(* IEC 61131-3 sources: plcassist-cli/packages/volt-lsp-iec/test-corpus/pro2193/Device/Plc Logic/Application/09 Misc/Library Manager/L_TT1P_TechnologyModules, 210 files *)

(* ---- L_MB1P_CONSTANTS.gvl ---- *)
VAR_GLOBAL
	GC_DWCHECKIDTAPPETREF : DWORD := 16#DC34;
	GC_LREPSILON : LREAL := 1E-06;
	GC_POSITIVE_LIMIT_32BIT : LREAL := 2147483647;
	GC_NEGATIVE_LIMIT_32BIT : LREAL := -2147483647;
	GC_PI : LREAL := 3.1415926535897931;
END_VAR

(* ---- L_MB1P_GLOBAL.gvl ---- *)
VAR_GLOBAL
END_VAR

(* ---- ITF_DATABUS.itf ---- *)
INTERFACE ITF_DATABUS
END_INTERFACE

(* ---- ITF_DATABUSPAR.itf ---- *)
INTERFACE ITF_DATABUSPAR
END_INTERFACE

(* ---- ITF_LIST.itf ---- *)
INTERFACE ITF_LIST
END_INTERFACE

(* ---- GETBOOLEANPROPERTY.fun ---- *)
FUNCTION GETBOOLEANPROPERTY : BOOL
VAR_INPUT
	STKEY : WSTRING;
END_VAR
END_FUNCTION

(* ---- GETCOMPANY.fun ---- *)
FUNCTION GETCOMPANY : WSTRING
END_FUNCTION

(* ---- GETNUMBERPROPERTY.fun ---- *)
FUNCTION GETNUMBERPROPERTY : DINT
VAR_INPUT
	STKEY : WSTRING;
END_VAR
END_FUNCTION

(* ---- GETTEXTPROPERTY.fun ---- *)
FUNCTION GETTEXTPROPERTY : WSTRING
VAR_INPUT
	STKEY : WSTRING;
END_VAR
END_FUNCTION

(* ---- GETTEXTPROPERTY2.fun ---- *)
FUNCTION GETTEXTPROPERTY2 : POINTER TO WSTRING
VAR_INPUT
	STKEY : WSTRING;
END_VAR
END_FUNCTION

(* ---- GETTITLE.fun ---- *)
FUNCTION GETTITLE : WSTRING
END_FUNCTION

(* ---- GETVERSION.fun ---- *)
FUNCTION GETVERSION : VERSION
END_FUNCTION

(* ---- GETVERSIONPROPERTY.fun ---- *)
FUNCTION GETVERSIONPROPERTY : VERSION
VAR_INPUT
	STKEY : WSTRING;
END_VAR
END_FUNCTION

(* ---- L_MB1P_CALCDISTBETWEEN3DPOINTS.fun ---- *)
FUNCTION L_MB1P_CALCDISTBETWEEN3DPOINTS : LREAL
VAR_INPUT
	LRX1 : LREAL;
	LRY1 : LREAL;
	LRZ1 : LREAL;
	LRX2 : LREAL;
	LRY2 : LREAL;
	LRZ2 : LREAL;
END_VAR
END_FUNCTION

(* ---- L_MB1P_CALCIDENDIAMETERBASE.fun ---- *)
FUNCTION L_MB1P_CALCIDENDIAMETERBASE : LREAL
VAR_IN_OUT
	LRLINEDIST : LREAL;
	LRDIAMCALCDIST : LREAL;
END_VAR
END_FUNCTION

(* ---- L_MB1P_CALCIDENDIAMETERSTATE.fun ---- *)
FUNCTION L_MB1P_CALCIDENDIAMETERSTATE : LREAL
VAR_IN_OUT
	LRDANCERPOSSTART : LREAL;
	LRDANCERPOSEND : LREAL;
	LRDIAMCALCDIST : LREAL;
	LRDANCERMATERIALLENGTH : LREAL;
END_VAR
END_FUNCTION

(* ---- L_MB1P_CHECK_CAMREFCHANGED.fun ---- *)
FUNCTION L_MB1P_CHECK_CAMREFCHANGED : BOOL
VAR_INPUT
	CAMREFNEW : MC_CAM_REF;
	CAMREFOLD : MC_CAM_REF;
END_VAR
END_FUNCTION

(* ---- L_MB1P_CHECK_CAMREFVALID.fun ---- *)
FUNCTION L_MB1P_CHECK_CAMREFVALID : BOOL
VAR_INPUT
	CAMREF : MC_CAM_REF;
END_VAR
END_FUNCTION

(* ---- L_MB1P_CHECKREQUESTSINFO.fun ---- *)
FUNCTION L_MB1P_CHECKREQUESTSINFO : BOOL
VAR_OUTPUT
	XRTRIG : BOOL;
	XFTRIG : BOOL;
	DWRTRIG : DWORD;
	DWFTRIG : DWORD;
END_VAR
VAR_IN_OUT
	DWREQUESTSINFO : DWORD;
	DWREQUESTSINFO_OLD : DWORD;
END_VAR
END_FUNCTION

(* ---- L_MB1P_CONVERTDWORDTOLREALMODULOPOS.fun ---- *)
FUNCTION L_MB1P_CONVERTDWORDTOLREALMODULOPOS : LREAL
VAR_INPUT
	DWIN : DWORD;
	LRPERIOD : LREAL;
END_VAR
END_FUNCTION

(* ---- L_MB1P_CONVERTLREALTODWORDLMODULOPOS.fun ---- *)
FUNCTION L_MB1P_CONVERTLREALTODWORDLMODULOPOS : DWORD
VAR_INPUT
	LRIN : LREAL;
	LRPERIOD : LREAL;
END_VAR
END_FUNCTION

(* ---- L_MB1P_CONVERTPOSTOMODULOPOS.fun ---- *)
FUNCTION L_MB1P_CONVERTPOSTOMODULOPOS : LREAL
VAR_INPUT
	LRPOS : LREAL;
	LRPERIOD : LREAL;
END_VAR
VAR_OUTPUT
	DIREVCOUNTER : DINT;
END_VAR
END_FUNCTION

(* ---- L_MB1P_CONVERTPOSTOMODULOPOSEXTENDED.fun ---- *)
FUNCTION L_MB1P_CONVERTPOSTOMODULOPOSEXTENDED : LREAL
VAR_INPUT
	LRPOS : LREAL;
	LRPERIOD : LREAL;
END_VAR
VAR_OUTPUT
	DIREVCOUNTER : DINT;
END_VAR
END_FUNCTION

(* ---- L_MB1P_CONVERTPOSTOMODULOPOSFMOD.fun ---- *)
FUNCTION L_MB1P_CONVERTPOSTOMODULOPOSFMOD : LREAL
VAR_INPUT
	LRPOS : LREAL;
	LRPERIOD : LREAL;
END_VAR
END_FUNCTION

(* ---- L_MB1P_DIV.fun ---- *)
FUNCTION L_MB1P_DIV : LREAL
VAR_INPUT
	A : LREAL;
	B : LREAL;
END_VAR
END_FUNCTION

(* ---- L_MB1P_GETOVERRIDEFADINGTIME.fun ---- *)
FUNCTION L_MB1P_GETOVERRIDEFADINGTIME : BOOL
VAR_IN_OUT
	AXESGROUP : AXES_GROUP_KIN;
	WNUMOFMOVEFBS : WORD;
	LROVERRIDEFADINGTIME : LREAL;
	LRMAXVEL : LREAL := 0;
	LRMAXACC : LREAL := 0;
	LRMAXDEC : LREAL := 0;
	LRMAXJERK : LREAL := 0;
END_VAR
END_FUNCTION

(* ---- L_MB1P_GETPROFILETIMEMOVECONTPATH.fun ---- *)
FUNCTION L_MB1P_GETPROFILETIMEMOVECONTPATH : LREAL
VAR_IN_OUT
	AXESGROUP : AXES_GROUP_KIN;
	FB_MOVECONTPATH : L_MC4P_MoveContPath;
END_VAR
END_FUNCTION

(* ---- L_MB1P_GETTASKCYCLE.fun ---- *)
FUNCTION L_MB1P_GETTASKCYCLE : LREAL
END_FUNCTION

(* ---- L_MB1P_HLPCALCKOEFPOLY5THORD.fun ---- *)
FUNCTION L_MB1P_HLPCALCKOEFPOLY5THORD : ARRAY [0..5] OF LREAL
VAR_INPUT
	LRYPOSSTART : LREAL;
	LRYVELSTART : LREAL;
	LRYACCSTART : LREAL;
	LRYPOSEND : LREAL;
	LRYVELEND : LREAL;
	LRYACCEND : LREAL;
END_VAR
VAR_OUTPUT
	ALRKOEF : ARRAY [0..5] OF LREAL;
END_VAR
END_FUNCTION

(* ---- L_MB1P_HLPCALCYOFPOLY5THORDBASE.fun ---- *)
FUNCTION L_MB1P_HLPCALCYOFPOLY5THORDBASE : LREAL
VAR_OUTPUT
	LRYPOSSCALED : LREAL;
END_VAR
VAR_IN_OUT
	LRXPOSSCALED : LREAL;
	ALRKOEF : ARRAY [0..5] OF LREAL;
END_VAR
END_FUNCTION

(* ---- L_MB1P_HLPCALCYOFPOLY5THORDSTATE.fun ---- *)
FUNCTION L_MB1P_HLPCALCYOFPOLY5THORDSTATE : LREAL
VAR_INPUT
	LRXPOSSTART : LREAL;
	LRXPOSEND : LREAL := 1;
	LRSETXPOS : LREAL;
	ALRKOEF : ARRAY [0..5] OF LREAL;
END_VAR
VAR_OUTPUT
	LRYPOSSCALED : LREAL;
END_VAR
END_FUNCTION

(* ---- L_MB1P_HLPCHECKDIRECTION.fun ---- *)
FUNCTION L_MB1P_HLPCHECKDIRECTION : INT
VAR_IN_OUT
	LRPOSFIFOX : ARRAY [1..20] OF LREAL;
	LRLEN : LREAL;
END_VAR
END_FUNCTION

(* ---- L_MB1P_HLPDELTAVELTIMEEXTENDED.fun ---- *)
FUNCTION L_MB1P_HLPDELTAVELTIMEEXTENDED : BOOL
VAR_INPUT
	LRVELSTART : LREAL;
	LRACCSTART : LREAL;
	LRMAXACC : LREAL;
	LRMAXJERK : LREAL;
END_VAR
VAR_OUTPUT
	LRTIME : LREAL;
	LRDIST : LREAL;
END_VAR
END_FUNCTION

(* ---- L_MB1P_HLPDELTAVELTIMESTATE.fun ---- *)
FUNCTION L_MB1P_HLPDELTAVELTIMESTATE : BOOL
VAR_INPUT
	LRVELSTART : LREAL;
	LRACCSTART : LREAL;
	LRVELTARGET : LREAL;
	LRACCTARGET : LREAL;
	LRMAXACC : LREAL;
	LRMAXDEC : LREAL;
	LRMAXJERK : LREAL;
END_VAR
VAR_OUTPUT
	LRTIME : LREAL;
	LRDIST : LREAL;
END_VAR
END_FUNCTION

(* ---- L_MB1P_HLPDELTAVELTIMETOCONTANTVEL.fun ---- *)
FUNCTION L_MB1P_HLPDELTAVELTIMETOCONTANTVEL : BOOL
VAR_INPUT
	LRACCSTART : LREAL;
	LRMAXJERK : LREAL;
	WMODE : WORD;
END_VAR
VAR_OUTPUT
	LRVEL : LREAL;
	LRTIME : LREAL;
	LRDIST : LREAL;
END_VAR
END_FUNCTION

(* ---- L_MB1P_HLPDYNAMIZE.fun ---- *)
FUNCTION L_MB1P_HLPDYNAMIZE : LREAL
VAR_INPUT
	LRDIFF : LREAL;
	LRTIME : LREAL;
	LRCYCLETIME : LREAL;
END_VAR
END_FUNCTION

(* ---- L_MB1P_HLPFITCYCLE.fun ---- *)
FUNCTION L_MB1P_HLPFITCYCLE : LREAL
VAR_INPUT
	LRPOS : LREAL;
	LRLEN : LREAL;
END_VAR
END_FUNCTION

(* ---- L_MB1P_HLPFITCYCLELIM.fun ---- *)
FUNCTION L_MB1P_HLPFITCYCLELIM : BOOL
VAR_INPUT
	PLRPOS : POINTER TO LREAL;
	LRLEN : LREAL;
END_VAR
END_FUNCTION

(* ---- L_MB1P_HLPGEARRES.fun ---- *)
FUNCTION L_MB1P_HLPGEARRES : LREAL
VAR_INPUT
	LRINPUT : LREAL;
	LRNUM : LREAL;
	LRDEN : LREAL;
END_VAR
END_FUNCTION

(* ---- L_MB1P_HLPISLIMITED.fun ---- *)
FUNCTION L_MB1P_HLPISLIMITED : BOOL
VAR_INPUT
	LRVAL : LREAL;
END_VAR
END_FUNCTION

(* ---- L_MB1P_HLPMODULOADD.fun ---- *)
FUNCTION L_MB1P_HLPMODULOADD : LREAL
VAR_INPUT
	LRINPUT : LREAL;
	LROFFSET : LREAL;
	LRLENGHT : LREAL;
END_VAR
END_FUNCTION

(* ---- L_MB1P_HLPMODULODIFF.fun ---- *)
FUNCTION L_MB1P_HLPMODULODIFF : LREAL
VAR_INPUT
	LRDIFF : LREAL;
	LRLEN : LREAL;
END_VAR
END_FUNCTION

(* ---- L_MB1P_HLPMODULOOFFSET.fun ---- *)
FUNCTION L_MB1P_HLPMODULOOFFSET : LREAL
VAR_INPUT
	LROFFSET : LREAL;
	LRLENGTH : LREAL;
	PLROFFSETBASE : POINTER TO LREAL;
END_VAR
END_FUNCTION

(* ---- L_MB1P_HLPMODULOSUB.fun ---- *)
FUNCTION L_MB1P_HLPMODULOSUB : LREAL
VAR_INPUT
	LRDIFF : LREAL;
	LRLEN : LREAL;
END_VAR
END_FUNCTION

(* ---- L_MB1P_HLPMODULOZEROPOS.fun ---- *)
FUNCTION L_MB1P_HLPMODULOZEROPOS : BOOL
VAR_INPUT
	PLRPOS : POINTER TO LREAL;
	LRLENINT : LREAL;
END_VAR
END_FUNCTION

(* ---- L_MB1P_HLPPOLY4RG.fun ---- *)
FUNCTION L_MB1P_HLPPOLY4RG : LREAL
VAR_INPUT
	LRX : LREAL;
END_VAR
END_FUNCTION

(* ---- L_MB1P_HLPPT1FILT.fun ---- *)
FUNCTION L_MB1P_HLPPT1FILT : LREAL
VAR_INPUT
	LRVALUE : LREAL;
	LRINPUT : LREAL;
	LRNEW_N : LREAL;
END_VAR
END_FUNCTION

(* ---- L_MB1P_HLPSIGNNE.fun ---- *)
FUNCTION L_MB1P_HLPSIGNNE : BOOL
VAR_INPUT
	A : LREAL;
	B : LREAL;
END_VAR
END_FUNCTION

(* ---- L_MB1P_IDENTMAXPOSSIBLEDIAMETER.fun ---- *)
FUNCTION L_MB1P_IDENTMAXPOSSIBLEDIAMETER : LREAL
VAR_INPUT
	WIDENTDIAMCALCCYCLES : WORD := 1;
END_VAR
VAR_IN_OUT
	LRACTDANCERPOSIN : LREAL;
	LRMAXDANCERPOS : LREAL;
	LRDANCERMATERIALLENGTH : LREAL;
	LRDIAMCALCDIST : LREAL;
END_VAR
END_FUNCTION

(* ---- L_MB1P_LREQ.fun ---- *)
FUNCTION L_MB1P_LREQ : BOOL
VAR_INPUT
	LRVALUE : LREAL;
	LRTARGET : LREAL;
END_VAR
END_FUNCTION

(* ---- L_MB1P_LRGE.fun ---- *)
FUNCTION L_MB1P_LRGE : BOOL
VAR_INPUT
	LRVALUE : LREAL;
	LRTARGET : LREAL;
END_VAR
END_FUNCTION

(* ---- L_MB1P_LRGT.fun ---- *)
FUNCTION L_MB1P_LRGT : BOOL
VAR_INPUT
	LRVALUE : LREAL;
	LRTARGET : LREAL;
END_VAR
END_FUNCTION

(* ---- L_MB1P_LRLE.fun ---- *)
FUNCTION L_MB1P_LRLE : BOOL
VAR_INPUT
	LRVALUE : LREAL;
	LRTARGET : LREAL;
END_VAR
END_FUNCTION

(* ---- L_MB1P_LRLT.fun ---- *)
FUNCTION L_MB1P_LRLT : BOOL
VAR_INPUT
	LRVALUE : LREAL;
	LRTARGET : LREAL;
END_VAR
END_FUNCTION

(* ---- L_MB1P_LRNE.fun ---- *)
FUNCTION L_MB1P_LRNE : BOOL
VAR_INPUT
	LRVALUE : LREAL;
	LRTARGET : LREAL;
END_VAR
END_FUNCTION

(* ---- L_MB1P_MODULOCYCLE.fun ---- *)
FUNCTION L_MB1P_MODULOCYCLE : LREAL
VAR_INPUT
	LRPOSIN : LREAL;
	LRPOSITIONPERIOD : LREAL;
END_VAR
END_FUNCTION

(* ---- L_MB1P_POSITIONINSIDEWINDOW.fun ---- *)
FUNCTION L_MB1P_POSITIONINSIDEWINDOW : BOOL
VAR_INPUT
	LRPOSIN : LREAL;
	LRLOWERWINDOW : LREAL;
	LRUPPERWINDOW : LREAL;
END_VAR
VAR_OUTPUT
	XERROR : BOOL := FALSE;
END_VAR
VAR_IN_OUT
	AXIS : AXIS_REF;
END_VAR
END_FUNCTION

(* ---- L_MB1P_PROFILETIMEVALID.fun ---- *)
FUNCTION L_MB1P_PROFILETIMEVALID : BOOL
VAR_IN_OUT
	LRPROFILETIME : LREAL;
END_VAR
END_FUNCTION

(* ---- L_TT1P_CALCSYNCTIME.fun ---- *)
FUNCTION L_TT1P_CALCSYNCTIME : BOOL
VAR_INPUT
	LRACTMATERIALVEL : LREAL;
	LRACCMAX : LREAL;
	LRJERKSTART : LREAL;
	LRJERKEND : LREAL;
END_VAR
VAR_OUTPUT
	LRACCTIME : LREAL;
	LRACCDIST : LREAL;
END_VAR
END_FUNCTION

(* ---- SB_CALCULATEPRODUCTERROR.fun ---- *)
FUNCTION SB_CALCULATEPRODUCTERROR : LREAL
VAR_INPUT
	LRPRODUCTTARGETCORRECTED : LREAL;
	LRMASTERPOSITIONATDETECTION : LREAL;
	LRCORRECTEDFACTORCOMPAREPOSITION : LREAL;
	BYNUMBEROFTARGETS : BYTE;
	LRMASTERCYCLELENGTH : LREAL;
END_VAR
END_FUNCTION

(* ---- _L_MB1A_ANALOGINTOSPEEDOUT.fb ---- *)
FUNCTION_BLOCK _L_MB1A_ANALOGINTOSPEEDOUT
VAR_INPUT
	WINPUT : WORD;
	WUPPERLIM : WORD := 16000;
	WLOWERLIM : WORD := 0;
	LRUPPERSPEEDLIM : LREAL := 1000.0;
	LRLOWERSPEEDLIM : LREAL := -1000.0;
	RFILTTIME : REAL := 0.01;
	LRACC : LREAL := 1000;
	LRDEC : LREAL := 1000;
	LRJERK : LREAL := 100000;
	XNEGATIVEDIRECTION : BOOL;
	LRDEADBANDWINDOW : LREAL := 10;
END_VAR
VAR_OUTPUT
	LRSETSPEEDOUT : LREAL;
END_VAR
VAR
	LRSPEEDSETPOINT : LREAL;
	L_MB1P_RAMPGENERATOR1 : L_MC1P_RampGenerator;
END_VAR
END_FUNCTION_BLOCK

(* ---- _L_MB1A_IOSELECTMASK.fb ---- *)
FUNCTION_BLOCK _L_MB1A_IOSELECTMASK
VAR_INPUT
	XENABLE : BOOL;
	WNUMOFMASK : WORD := 3;
	XSELECTMASK : BOOL;
	XIP1 : BOOL;
	XIP2 : BOOL;
	XIP3 : BOOL;
	XIP4 : BOOL;
	XIP5 : BOOL;
	XIP6 : BOOL;
	XIP7 : BOOL;
	XIP8 : BOOL;
END_VAR
VAR_OUTPUT
	XBLINKEROUT : BOOL;
	WNOOUT : WORD;
	WMASK : WORD;
	AXOP1 : ARRAY [1..10] OF BOOL;
	AXOP2 : ARRAY [1..10] OF BOOL;
	AXOP3 : ARRAY [1..10] OF BOOL;
	AXOP4 : ARRAY [1..10] OF BOOL;
	AXOP5 : ARRAY [1..10] OF BOOL;
	AXOP6 : ARRAY [1..10] OF BOOL;
	AXOP7 : ARRAY [1..10] OF BOOL;
	AXOP8 : ARRAY [1..10] OF BOOL;
END_VAR
VAR
	XSELECTMASK_OLD : BOOL;
	XBLINKEROUT_OLD : BOOL;
	TON_1 : TON;
	TOF_1 : TOF := STRUCT(PT := TIME#400ms);
	WCNTR : WORD;
	XBLINKER : BOOL;
	XIP1_OLD : BOOL;
	XIP2_OLD : BOOL;
	XIP3_OLD : BOOL;
	XIP4_OLD : BOOL;
	XIP5_OLD : BOOL;
	XIP6_OLD : BOOL;
	XIP7_OLD : BOOL;
	XIP8_OLD : BOOL;
END_VAR
END_FUNCTION_BLOCK

METHOD CALL_BLINKER
END_METHOD

(* ---- _L_MB1P_ANALOGINPUTSPEEDCTRL.fb ---- *)
FUNCTION_BLOCK _L_MB1P_ANALOGINPUTSPEEDCTRL
VAR_INPUT
	WINPUT : WORD;
	WUPPERLIM : WORD := 10000;
	WLOWERLIM : WORD := 0;
	LRUPPERSPEEDLIM : LREAL := 1000;
	LRLOWERSPEEDLIM : LREAL := 0;
	LRDEADBAND : LREAL := 5;
	RFILTTIME : REAL := 0.01;
	LRACC : LREAL := 1000;
	LRDEC : LREAL := 1000;
	LRJERK : LREAL := 100000;
	XNEGATIVEDIRECTION : BOOL;
END_VAR
VAR_OUTPUT
	LRSETSPEEDOUT : LREAL;
END_VAR
VAR
	LRINPUTSCALED : LREAL;
	LRSPEEDSETPOINT : LREAL;
	L_D94A_FILTER : L_USPP_PT1Filter;
	L_MB1P_RAMPGENERATOR1 : L_MC1P_RampGenerator;
END_VAR
END_FUNCTION_BLOCK

(* ---- _L_MB1P_AXISCONTROLBYPOS.fb ---- *)
FUNCTION_BLOCK _L_MB1P_AXISCONTROLBYPOS
VAR_INPUT
	XENABLE : BOOL;
	LRSETPOSITION : LREAL;
	LRSETVELOCITY : LREAL;
	LRSETACCELERATION : LREAL;
	ESETVALUEMODE : L_MC1P_SetValueMode := L_MC1P_SetValueMode.Pos;
END_VAR
VAR_OUTPUT
	XBUSY : BOOL;
	XCOMMANDABORTED : BOOL;
	XERROR : BOOL;
	EERRORID : L_IE1P_Error;
	LRSETPOSOUT : LREAL;
END_VAR
VAR_IN_OUT
	AXIS : AXIS_REF;
END_VAR
VAR
	LRSETPOSITION_INT : LREAL;
	XENABLE_OLD : BOOL;
	XBUSY_OLD : BOOL;
	ESTATE : L_MB1P_States;
	MC_HALT1 : MC_HALT;
	FB_FOLLOWSETVALUES : L_MC1P_FollowSetValues;
END_VAR
END_FUNCTION_BLOCK

METHOD CALL_ERRORHANDLER
END_METHOD

METHOD CALL_FBMETHODS
END_METHOD

METHOD CALL_FB_FOLLOWSETVALUES
END_METHOD

METHOD CALL_MC_HALT
END_METHOD

METHOD CALL_MC_HALT_INPUT
END_METHOD

METHOD CALL_OUTPUT
END_METHOD

METHOD CALL_RESETCOMMANDS
END_METHOD

METHOD CALL_RESETOUTPUT
END_METHOD

METHOD CALL_STATEMACHINE
END_METHOD

METHOD CALL_S000_CYCLIC
END_METHOD

METHOD CALL_S001_INIT
END_METHOD

METHOD CALL_S002_READY
END_METHOD

METHOD CALL_S999_ERROR
END_METHOD

(* ---- _L_MB1P_AXISCONTROLBYVEL.fb ---- *)
FUNCTION_BLOCK _L_MB1P_AXISCONTROLBYVEL
VAR_INPUT
	XENABLE : BOOL;
	LRSETVELOCITY : LREAL;
END_VAR
VAR_OUTPUT
	XBUSY : BOOL;
	XCOMMANDABORTED : BOOL;
	XERROR : BOOL;
	EERRORID : L_IE1P_Error;
	LRSETVELOUT : LREAL;
END_VAR
VAR_IN_OUT
	AXIS : AXIS_REF;
END_VAR
VAR
	LRSETVELOCITY_INT : LREAL;
	XENABLE_OLD : BOOL;
	XBUSY_OLD : BOOL;
	ESTATE : L_MB1P_States;
	MC_HALT1 : MC_HALT;
	FB_FOLLOWSETVALUES : L_MC1P_FollowSetValues;
END_VAR
END_FUNCTION_BLOCK

METHOD CALL_ERRORHANDLER
END_METHOD

METHOD CALL_FBMETHODS
END_METHOD

METHOD CALL_FB_FOLLOWSETVALUES
END_METHOD

METHOD CALL_MC_HALT
END_METHOD

METHOD CALL_MC_HALT_INPUT
END_METHOD

METHOD CALL_OUTPUT
END_METHOD

METHOD CALL_RESETCOMMANDS
END_METHOD

METHOD CALL_RESETOUTPUT
END_METHOD

METHOD CALL_STATEMACHINE
END_METHOD

METHOD CALL_S000_CYCLIC
END_METHOD

METHOD CALL_S001_INIT
END_METHOD

METHOD CALL_S002_READY
END_METHOD

METHOD CALL_S999_ERROR
END_METHOD

(* ---- _TM_BASE.fb ---- *)
FUNCTION_BLOCK _TM_BASE
VAR
	DWVERSION : DWORD;
	DWID : DWORD;
	DWVENDORID : DWORD;
	BYCOUNTER : BYTE;
	XHARDWARECHECKPASSED : BOOL;
	XSYSTEMFAULT : BOOL;
END_VAR
END_FUNCTION_BLOCK

(* ---- _TM_BASICMOTIONBASE.fb ---- *)
FUNCTION_BLOCK _TM_BASICMOTIONBASE EXTENDS _TM_MotionControl
VAR_OUTPUT
	PPAR : POINTER TO _scPar_TM_BasicMotionHigh;
	PSF : POINTER TO _scSF_TM_BasicMotionHigh;
	PAP : POINTER TO _scAP_TM_BasicMotionHigh;
END_VAR
VAR_IN_OUT
	AXIS : AXIS_REF;
	XMOVEVELEXECUTE : BOOL;
	XMOVEABSEXECUTE : BOOL;
	XMOVERELEXECUTE : BOOL;
	LRSETPOS_DIST : LREAL;
	XDISABLESWLIMIT : BOOL;
	LROVERRIDE : LREAL;
	LROVERRIDEACC : LREAL;
	LROVERRIDEJERK : LREAL;
	XAXISREADY : BOOL;
	XCOMMANDABORTED : BOOL;
	XINPOSITION : BOOL;
	XHWLIMITSWITCHNEG : BOOL;
	XHWLIMITSWITCHPOS : BOOL;
	XSWLIMITENABLED : BOOL;
	XSWLIMITSWITCHNEG : BOOL;
	XSWLIMITSWITCHPOS : BOOL;
	EAXISSTATE : L_MC1P_AXIS_STATE;
	ECONTROLMODE : L_MC1P_ControlMode;
	LRACTVEL : LREAL;
	LRACTPOS : LREAL;
	LRSETPOSOUT : LREAL;
	LRSETVELOUT : LREAL;
	LRACTFOLLOWINGERROR : LREAL;
	XCONSTANTVELOCITY : BOOL;
	XACCELERATING : BOOL;
	XDECELERATING : BOOL;
	XDIRECTIONPOSITIVE : BOOL;
	XDIRECTIONNEGATIVE : BOOL;
END_VAR
VAR
	SCPAR_INT : _scPar_TM_BasicMotionHigh;
	XMOVEVELEXECUTE_INT : BOOL;
	XMOVEABSEXECUTE_INT : BOOL;
	XMOVERELEXECUTE_INT : BOOL;
	LRSETPOS_DIST_INT : LREAL;
	XDISABLESWLIMIT_INT : BOOL;
	LROVERRIDE_INT : LREAL := 1.0;
	LROVERRIDEACC_INT : LREAL := 1.0;
	LROVERRIDEJERK_INT : LREAL := 1.0;
	XCOMMANDABORTED_INT : BOOL;
END_VAR
END_FUNCTION_BLOCK

METHOD CALL_ABC
END_METHOD

METHOD CALL_ABC_INPUT
END_METHOD

METHOD CALL_ALLOCPOINTADR
END_METHOD

METHOD CALL_CTRLREQACTIVE : BOOL
END_METHOD

METHOD CALL_ERRORHANDLER
END_METHOD

METHOD CALL_FBMETHODS
END_METHOD

METHOD CALL_INITDONE
END_METHOD

METHOD CALL_INITROUTINE
END_METHOD

METHOD CALL_INTERNALCTRL
END_METHOD

METHOD CALL_OUTPUT
END_METHOD

METHOD CALL_OUTPUT_SF
END_METHOD

METHOD CALL_REQUESTS_EXT
END_METHOD

METHOD CALL_RESETCOMMANDS
END_METHOD

METHOD CALL_RESETOUTPUT
END_METHOD

METHOD CALL_STATEMACHINE
END_METHOD

METHOD CALL_S003_HOMING
END_METHOD

METHOD CALL_S013_MOVEVEL
END_METHOD

METHOD CALL_S014_MOVEABS
END_METHOD

METHOD CALL_S015_MOVEREL
END_METHOD

METHOD CALL_S017_EXTERNAL
END_METHOD

METHOD CALL_S995_HALT
END_METHOD

METHOD CALL_T000_ALLSTATES
END_METHOD

METHOD CALL_T002_READY
END_METHOD

(* ---- _TM_CROSSCUTTERBASE.fb ---- *)
FUNCTION_BLOCK _TM_CROSSCUTTERBASE EXTENDS _TM_MotionControl
VAR_OUTPUT
	PAP : POINTER TO _scAP_TM_CrossCutterHigh;
	PSF : POINTER TO _scSF_TM_CrossCutterHigh;
	PPAR : POINTER TO _scPar_TM_CrossCutterHigh;
	PPARBASE : POINTER TO _scPar_TM_CrossCutterBaseExtension;
END_VAR
VAR_IN_OUT
	MASTERAXIS : AXIS_REF;
	SLAVEAXIS : AXIS_REF;
	XEXECUTEMOVETOPARKPOS : BOOL;
	XSYNCCROSSCUTTER : BOOL;
	XSYNCOUTINSTANT : BOOL;
	XHOLDINPARKPOS : BOOL;
	LRPRODUCTLENGTH : LREAL;
	LRSETOVERSPEEDSCALED : LREAL;
	LRSETOFFSETMASTER : LREAL;
	XTRIMPOS : BOOL;
	XTRIMNEG : BOOL;
	XRESETTRIMOFFSET : BOOL;
	XINPARKPOS : BOOL;
	XSYNCHRONISED : BOOL;
	XACCDECSYNC : BOOL;
	XHOLDINPARKPOSACTIVE : BOOL;
	XCUTTINGACTIVE : BOOL;
	XCUTDONE : BOOL;
	LRACTCUTLENGTH : LREAL;
	BYSETTOOLNOOUT : BYTE;
	BYSETAREAOUT : BYTE;
	LROFFSET : LREAL;
	LROFFSETTRIM : LREAL;
	LROFFSETTOTAL : LREAL;
	LRSETXPOSOUT : LREAL;
	LRSETXVELOUT : LREAL;
	LRSETXACCOUT : LREAL;
	LRACTSLAVEFOLLOWINGERROR : LREAL;
	LRACTSLAVEPOS : LREAL;
	LRACTSLAVEVEL : LREAL;
	LRSLAVEMAXVEL : LREAL;
	LRSLAVEMAXACC : LREAL;
END_VAR
VAR
	XEXECUTEMOVETOPARKPOS_INT : BOOL;
	XSYNCCROSSCUTTER_INT : BOOL;
	XSYNCOUTINSTANT_INT : BOOL;
	XHOLDINPARKPOS_INT : BOOL;
	PMASTERAXIS : POINTER TO _AXIS_REF_REAL;
	LRPRODUCTLENGTH_INT : LREAL;
	LRSETOVERSPEEDSCALED_INT : LREAL;
	LRCUTTINGANGLE_INT : LREAL;
	LRSETOFFSETMASTER_INT : LREAL;
	LRSETOFFSETSLAVE_INT : LREAL;
	XTRIMPOS_INT : BOOL;
	XTRIMNEG_INT : BOOL;
	XRESETTRIMOFFSET_INT : BOOL;
	SCPAR_INT : _scPar_TM_CrossCutterHigh;
	SCPARBASE_INT : _scPar_TM_CrossCutterBaseExtension;
	LRSLAVEMAXVEL_INT : LREAL;
	LRSLAVEMAXACC_INT : LREAL;
	XHOMEEXECUTE_OLD : BOOL;
	LRMASTERVEL : LREAL;
	LRMASTERVEL_OLD : LREAL;
	LRMASTERVEL_OLD2 : LREAL;
	LRMASTERPOS_OLD : LREAL;
	LRACTMASTERPOS_OLD : LREAL;
	XMASTERAXISENABLED : BOOL;
	XMASTERAXISENABLED_OLD : BOOL;
	XCUTTINGACTIVE_OLD : BOOL;
	XRESETTRIMOFFSET_OLD : BOOL;
	XMASTERISSTANDSTILL : BOOL;
	XNEXTTOOLDIRECTIONPOSITIV : BOOL := TRUE;
	ECUTTINGPROCESSSTATE : L_TT1P_States := L_TT1P_States.INIT;
	BYPOSITIONINGSTATE : BYTE := 0;
	BYMASTEROFFSETSTEPPER : BYTE := 0;
	BYTOOLCIRCARRAYPREPARED : BYTE;
	XMASTERIS_FREEENCODER : BOOL;
	XEXECUTETRANSITIONCYCLES : BOOL;
	XINVALIDCROSSCUTTERPARAMETRS : BOOL;
	XINVALIDCUTTINGPARAMETRS : BOOL;
	XMASTERNOTROTATIVE : BOOL;
	XWARNINGINVALIDPRODUCTLENGTH : BOOL;
	XINVALIDPRODUCTLENGTH : BOOL;
	XINVALIDCUTTINGANGLE : BOOL;
	XSLAVEOUTOFSCALE : BOOL;
	XMASTEROUTOFSCALE : BOOL;
	XSLAVERECEIVEDGAPS : BOOL;
	XINVALIDCAMSELECTED : BOOL;
	XWARNINGINVALIDCAMSELECTED : BOOL;
	ILOOPCNTR : INT;
	UIVARTEMP : UINT;
	IVARTEMP : INT;
	LRVARTEMP : LREAL;
	LRVARTEMP2 : LREAL;
	LRVARTEMP3 : LREAL;
	LRVARTEMP4 : LREAL;
	LRTEMPSTOPLENGTH : LREAL;
	LRTEMPSTARTLENGTH : LREAL;
	LRXDISTINPARKPOS : LREAL;
	XXPOSSYNCRONISEDMASTERPOS : BOOL;
	XCUTTINGPARISCHANGED : BOOL;
	XCAMDIRECTCHANGE_LOCK : BOOL;
	LRSETMASTERTRIMOFFSET_INT : LREAL;
	LRSETOFFSETMASTER_LOCK : LREAL;
	LRSETMASTERTRIMOFFSET_LOCK : LREAL;
	LRSETMASTERTRIMOFFSET_SAVE : LREAL;
	LRACTMASTERPOSSTART : LREAL;
	IMASTERPERIODCNT : INT;
	LRLENGTHCALCULATOR : LREAL;
	LROVERSPEEDUPPERLIMIT : LREAL := 2;
	ECUTTINGMODE_LOCK : L_TT1P_CuttingModeState;
	BYCAMCONTINUOUSNO_LOCK : BYTE := 1;
	BYNUMOFTOOLS_LOCK : BYTE;
	LRPRODUCTLENGTH_LOCK : LREAL;
	LRPRODUCTLENGTH_LOCK_OLD : LREAL;
	LRCUTLENGTH_LOCK : LREAL;
	LROSCILLATION_LOCK : LREAL := 0;
	LRSETOVERSPEEDSCALED_LOCK : LREAL;
	LROVERSPEEDFACTOR_LOCK : LREAL;
	LROVERSPEEDFACTOR_LOCK_OLD : LREAL;
	LRCUTTINGANGLE_LOCK : LREAL;
	LRSCALINGMASTER_LOCK : LREAL := 1;
	LRTOOLTOOLDIST_LOCK : LREAL;
	LRTOOLTOOLCIRCUMFERENCEDIST_LOCK : LREAL;
	LRCIRCUMFERENCE_LOCK : LREAL;
	LRCIRCUMFERENCEINV_LOCK : LREAL;
	XHOLDINPARKPOS_LOCK : BOOL;
	LRFACTOR_ANGLETOSLAVEUNITS_LOCK : LREAL;
	LRFACTOR_ANGLETOMASTERUNITS_LOCK : LREAL;
	LRFACTOR_SLAVEUNITSTOMASTERUNITS_LOCK : LREAL;
	LRFACTOR_MASTERUNITSTOSLAVEUNITS_LOCK : LREAL;
	LRFACTOR_PRODUCTUNITSTOMASTERUNITS_LOCK : LREAL;
	LRFACTOR_PRODUCTUNITSTOMASTERUNITSINV_LOCK : LREAL;
	LRFACTOR_PRODUCTUNITSTOMASTERUNITSINV_OLD : LREAL;
	XFIRSTCUT : BOOL;
	XCONTINUOUSMODE : BOOL := TRUE;
	BYSETCAMTABLENO : BYTE;
	BYREQUESTSSETCAMTABLE : BYTE;
	BYREQUESTSSETCAMTABLE_OLD : BYTE;
	SCSYNCSTARTLENGTH : L_MC2P_CamDataXYVA;
	SCSYNCSTOPLENGTH : L_MC2P_CamDataXYVA;
	SCASYNCLENGTH : L_MC2P_CamDataXYVA;
	SCSTARTLENGTH : L_MC2P_CamDataXYVA;
	SCSTOPLENGTH : L_MC2P_CamDataXYVA;
	LRSTANDSTILLLENGTH : LREAL;
	LRY_START : LREAL := 0;
	LRY_PARK : LREAL := 180;
	LRY_END : LREAL := 360;
	LRX_START : LREAL := 0;
	LRX_ENDSYNCPOS : LREAL := 10;
	LRX_STARTPARKPOS : LREAL := 180;
	LRX_ENDPARKPOS : LREAL := 180;
	LRX_STARTSYNCPOS : LREAL := 350;
	LRX_END : LREAL := 360;
	LRY_END_PREVIOUSLY : LREAL := 360;
	LRY_CUTLENGTHCALCULATOR : LREAL := 360;
	LRSETOVERSPEEDSCALED_LOCK_PREVIOUSLY : LREAL;
	FM_CAMCREATOR_START : L_MB1P_CamCreator;
	FM_CAMCREATOR_STOP : L_MB1P_CamCreator;
	FM_CAMCREATOR_CONTINUOUS : ARRAY [1..2] OF L_MB1P_CamCreator;
	FM_CAMCREATOR_STANDSTILL : L_MB1P_CamCreator;
	CAM_START_P : ARRAY [0..3] OF L_MC2P_CamDataXYVA;
	CAM_STOP_P : ARRAY [0..3] OF L_MC2P_CamDataXYVA;
	CAM_CONTINUOUS_P : ARRAY [1..2] OF ARRAY [0..3] OF L_MC2P_CamDataXYVA;
	CAM_STOPSTART_P : ARRAY [1..2] OF ARRAY [0..5] OF L_MC2P_CamDataXYVA;
	CAM_STANDSTILL_P : ARRAY [0..1] OF L_MC2P_CamDataXYVA;
	CAMTABLEATFLEXCAM : MC_CAM_REF;
	LRYOFFSET : LREAL;
	LRENDOFPROFILEWINDOWSIZE : LREAL := 0;
	_FC_XMASTERABSOLUTE : BOOL;
	_FC_XSLAVEABSOLUTE : BOOL;
	_FC_XPERIODIC : BOOL;
	_FC_XTRIMMASTERNEG : BOOL;
	_FC_XTRIMMASTERPOS : BOOL;
	_FC_LRSETOFFSETMASTER : LREAL;
	_FC_LRSETOFFSETSLAVE : LREAL;
	_FC_EPOSCTRLDIRECTION : L_MC2P.L_MC2P_ReverseCtrlDirection;
	_FC_EOFFSETMODEMASTER : L_MC2P.L_MC2P_OffsetMode;
	_FC_EOFFSETMODESLAVE : L_MC2P.L_MC2P_OffsetMode;
	_FC_XHOLDPROFGENMASTER : BOOL;
	_FC_ESYNCMODE : L_MC2P.L_MC2P_ClutchMode;
	_FC_ESYNCDIRECTION : L_MC2P.L_MC2P_ClutchDirection;
	_FC_LRMASTERSYNCINDIST : LREAL;
	_FC_LRMASTERSYNCINPOS : LREAL;
	_FC_LRMASTERSYNCOUTDIST : LREAL;
	_FC_LRSLAVESYNCOUTPOS : LREAL;
	_FC_LRSYNCINTIME : LREAL;
	_FC_LRSYNCOUTTIME : LREAL;
	_FC_LRSYNCOUTINSTANTDEC : LREAL;
	_FC_XENABLE : BOOL;
	_FC_XSYNCPOS : BOOL;
	_FC_XSYNCCAM : BOOL;
	_FC_XDIRECTCHANGE : BOOL;
	_FC_XSYNCOUTINSTANT : BOOL;
	_FC_LRSYNCCAMVEL : LREAL;
	_FC_LRSYNCCAMACC : LREAL;
	_FC_LRSYNCCAMDEC : LREAL;
	_FC_LRSYNCCAMJERK : LREAL;
	_FC_LRSETXPOSOUT : LREAL;
	_FC_LRSETXVELOUT : LREAL;
	_FC_LRSETXACCOUT : LREAL;
	_FC_LRSETYPOSOUT : LREAL;
	_FC_LRSETYVELOUT : LREAL;
	_FC_LRSETYACCOUT : LREAL;
	_FC_LRSETSLAVEPOSOUT : LREAL;
	_FC_LRSETSLAVEVELOUT : LREAL;
	_FC_LRSETSLAVEACCOUT : LREAL;
	_FC_XENDOFPROFILE : BOOL;
	_FC_XACCDECSYNC : BOOL;
	_FC_XSYNCHRONISED : BOOL;
	_FC_LRSETOFFSETMASTEROUT : LREAL;
	_FC_XENDOFCYCLE : BOOL;
	_FC_LRSETXPOS : LREAL;
	_FC_XCAMSYNCHRONISED : BOOL;
	_FC_XDONE : BOOL;
	_FC_XBUSY : BOOL;
	_FC_LRSETMASTERTRIMOFFSETOUT : LREAL;
	_FC_XENDOFPROFNEGATIVE : BOOL;
	_FC_LWENDOFPROFILECHECKSUM : LWORD;
	FM_FLEXCAMHIGH : L_MC2P_FlexCamHigh;
	FB_CONTROLSETVALUES : L_MC1P_ControlSetValues;
	L_MB1P_DIFFERENTIATE1 : L_MC2P_Differentiate;
	XINTERNALERROR : BOOL;
	WINTERNALERRORID : WORD;
	LWTCHECKSUM_INT : LWORD;
END_VAR
END_FUNCTION_BLOCK

METHOD CALL_ALLOCPOINTADR
END_METHOD

METHOD CALL_CTRLREQACTIVE : BOOL
END_METHOD

METHOD CALL_ERRORHANDLER
END_METHOD

METHOD CALL_ERRORHANDLER_STATECUTTING
END_METHOD

METHOD CALL_FBMETHODS
END_METHOD

METHOD CALL_FBMETHODS_BEFOREFLEXCAM
END_METHOD

METHOD CALL_FB_CONTROLAXISBYPOS
END_METHOD

METHOD CALL_FB_DIFFERENTIATEPOSITION
END_METHOD

METHOD CALL_FM_CAMCREATOR_CONTINUOUS1
END_METHOD

METHOD CALL_FM_CAMCREATOR_CONTINUOUS2
END_METHOD

METHOD CALL_FM_CAMCREATOR_START
END_METHOD

METHOD CALL_FM_CAMCREATORS
END_METHOD

METHOD CALL_FM_FLEXCAM
END_METHOD

METHOD CALL_FM_FLEXCAM_INPUT
END_METHOD

METHOD CALL_INITDONE
END_METHOD

METHOD CALL_INITROUTINE
END_METHOD

METHOD CALL_INTERNALCTRL
END_METHOD

METHOD CALL_INTERNALCTRLBASEEXTENSION
END_METHOD

METHOD CALL_MASTEROFFSET
END_METHOD

METHOD CALL_MASTERTRIMM
END_METHOD

METHOD CALL_OUTPUT
END_METHOD

METHOD CALL_OUTPUTMINMAXVALUES
END_METHOD

METHOD CALL_OUTPUT_SF
END_METHOD

METHOD CALL_PARSYNCINCAM
END_METHOD

METHOD CALL_PARSYNCOUT
END_METHOD

METHOD CALL_REQUESTSSETCAMTABLE
END_METHOD

METHOD CALL_REQUESTSSETCAMTABLECTRL
END_METHOD

METHOD CALL_REQUESTS_EXT
END_METHOD

METHOD CALL_RESETCOMMANDS
END_METHOD

METHOD CALL_RESETOUTPUT
END_METHOD

METHOD CALL_SETTOOLNOOUT
END_METHOD

METHOD CALL_STATEMACHINE
END_METHOD

METHOD CALL_ABC
END_METHOD

METHOD CALL_CALCACTXKOORDINATEN
END_METHOD

METHOD CALL_CALCCAM_CONTINUOUS
END_METHOD

METHOD CALL_CALCCAM_START
END_METHOD

METHOD CALL_CALCSYNCARRAY
END_METHOD

METHOD CALL_CHECKCUTTINGPARCHANGES
END_METHOD

METHOD CALL_CONTINUOUSCAMSETYOFFSET
END_METHOD

METHOD CALL_CUTLENGTHCALCULATOR
END_METHOD

METHOD CALL_INIT_FLEXCAM
END_METHOD

METHOD CALL_LOCKCAMTABLE
END_METHOD

METHOD CALL_LOCKCROSSCUTTERPAR
END_METHOD

METHOD CALL_LOCKCUTTINGPAR
END_METHOD

METHOD CALL_LOCKCUTTINGPAR_ECCMODE_0
END_METHOD

METHOD CALL_LOCKCUTTINGPAR_ECCMODE_1
END_METHOD

METHOD CALL_PREPARENEXTCUT
END_METHOD

METHOD CALL_PREPARENEXTCUT_ECCMODEPAR
END_METHOD

METHOD CALL_RESETALLCAMCREATOR
END_METHOD

METHOD CALL_SEARCHACTYCOORDINATE
END_METHOD

METHOD CALL_SEARCHPARKPOS
END_METHOD

METHOD CALL_SETNEXTCAMCREATOR_CONTINUOUS
END_METHOD

METHOD CALL_YCOORDINATEMANAGER
END_METHOD

METHOD CALL_CP_000_CYCLIC
END_METHOD

METHOD CALL_CP_001_INIT
END_METHOD

METHOD CALL_CP_001_INIT_OLD
END_METHOD

METHOD CALL_CP_141_IN_PARK_POS
END_METHOD

METHOD CALL_CP_142_ASYNC_PHASE
END_METHOD

METHOD CALL_CP_143_ENTRY_IN_SYNC_PHASE
END_METHOD

METHOD CALL_CP_143_ENTRY_IN_SYNC_PHASE_TRANSITION
END_METHOD

METHOD CALL_CP_144_EXIT_SYNC_PHASE
END_METHOD

METHOD CALL_CP_144_EXIT_SYNC_PHASE_TRANSITION
END_METHOD

METHOD CALL_CP_145_CLUTCH_CLOSE
END_METHOD

METHOD CALL_CP_146_CLUTCH_OPEN
END_METHOD

METHOD CALL_CP_148_HOLD_IN_PARK_POS
END_METHOD

METHOD CALL_CP_148_HOLD_IN_PARK_POS_CONTINUECUTTING
END_METHOD

METHOD CALL_CP_148_HOLD_IN_PARK_POS_ENDOFPROFILE
END_METHOD

METHOD CALL_CP_802_STOP_IN_PARK_POS
END_METHOD

METHOD CALL_CP_900_DONE
END_METHOD

METHOD CALL_CUTTING_PROCESS
END_METHOD

METHOD CALL_S000_CYCLIC
END_METHOD

METHOD CALL_S002_READY
END_METHOD

METHOD CALL_S030_SYNCHRONISING_POS
END_METHOD

METHOD CALL_S030_SYNCHRONISING_POS_ECCMODESELECT
END_METHOD

METHOD CALL_S030_SYNCHRONISING_POS_ECCMODE_0
END_METHOD

METHOD CALL_S030_SYNCHRONISING_POS_ECCMODE_1
END_METHOD

METHOD CALL_S032_POSITIONING_TO_START_POS
END_METHOD

METHOD CALL_S034_POSITIONING_TO_PARK_POS
END_METHOD

METHOD CALL_S035_CUTTING
END_METHOD

METHOD CALL_S996_STOP
END_METHOD

METHOD CALL_S999_ERROR
END_METHOD

METHOD CALL_T002_READY
END_METHOD

(* ---- _TM_CROSSCUTTERSTATE.fb ---- *)
FUNCTION_BLOCK _TM_CROSSCUTTERSTATE EXTENDS _TM_CrossCutterBase
VAR_IN_OUT
	XTEACHMARKWINDOW : BOOL;
	XMARKRECEIVE : BOOL;
	LRACTMARKPOSIN : LREAL;
	LRCYCPOSEXTENCODER : LREAL;
	XGEARFACTORCORR : BOOL;
	XGEARFACTORCORRHOLD : BOOL;
	XTRQCTRLACTIVE : BOOL;
	LRSETMOTORPRECTRLTRQOUT : LREAL;
	XREGISTERCTRLACTIVE : BOOL;
	XTEACHMARKWINDOWACTIVE : BOOL;
	LRSETREGPOSOUT : LREAL;
	LRMARKSENSORPOS : LREAL;
	LRREGMARKPOS : LREAL;
	LRACTMARKERROR : LREAL;
	LRACTMARKDIST : LREAL;
	XMARKRECEIVED : BOOL;
	XCORRACTIVE : BOOL;
	XCORRLIMITED : BOOL;
	XMARKWINDOWOPEN : BOOL;
	XMARKOUTOFWINDOW : BOOL;
	XMARKNOTDETECTED : BOOL;
	XMARKWINDOWTEACHED : BOOL;
	XLOADREGPOS : BOOL;
	LRLOADREGPOS : LREAL;
	LRAVERAGEGEARFACTORCORR : LREAL;
	XGEARFACTORCORRLIMITED : BOOL;
END_VAR
VAR
	XTEACHMARKWINDOW_INT : BOOL;
	XGEARFACTORCORR_INT : BOOL;
	XGEARFACTORCORRHOLD_INT : BOOL;
	LRCYCMASTERPOS_INT : LREAL;
	XLOADREGPOS_INT : BOOL;
	LRLOADREGPOS_INT : LREAL;
	XMARKRECEIVED_OLD : BOOL;
	XTEACHMARKWINDOW_OLD : BOOL;
	XLOADREGPOS_OLD : BOOL;
	AP11_XSETCUTLENGTHINPRODUCT_OLD : BOOL;
	EWARNINGID : WORD;
	FM_REGISTERCONTROLSTATE_LRACTVEL_OLD : LREAL;
	DNNUMAXISY_INT : DWORD := 1;
	DNDENAXISY_INT : DWORD := 1;
	LRCYCLELENGTHEXTENCODER : LREAL;
	XINVALIDCUTPRODUCTFORMAT : BOOL;
	XSCSCALINGVALID : BOOL := FALSE;
	XENABLETORQUEFOLLOWER : BOOL;
	XENABLEREGCTRLCORR : BOOL;
	XINVALIDTEACHMARKPOS : BOOL;
	LRCYCPOSEXTENCODER_OLD : LREAL;
	XWARNINGINVALIDMARKRECIVED : BOOL;
	XTAKENEXTSTACKPOS : BOOL;
	LRSTACKLATESTDIST : LREAL;
	ETPMODE_LOCK : L_TT1P_TpMode := L_TT1P_TpMode.TpFromMaster;
	LRSENSORTOOLDIST_LOCK : LREAL;
	LRMARKPOS_LOCK : LREAL;
	XFIRSTCUTOFARRAY : BOOL;
	XCUTLENGTHINPRODUCTCHANGED_LOCK : BOOL;
	ISETNOCUTLENGTH_LOCK : INT;
	ISETNOOFMAXCUTLENGTH_LOCK : INT;
	LRUPPERCORRPOS_LOCK : LREAL;
	LRLOWERCORRPOS_LOCK : LREAL;
	ALRCUTLENGTHINPRODUCT_LOCK : ARRAY [1..10] OF LREAL;
	LRMARKSENSORPOS_LOCK : LREAL;
	LRREGISTERLENGTH_LOCK : LREAL;
	LRMINLOWERCORRPOS : LREAL;
	XCORRINSAMECYCLE : BOOL;
	LRFACTOR_NMOTOR_D_NAPPL : LREAL := 1;
	LRFACTOR_NAPPL_D_NMOTOR : LREAL := 1;
	LRFACTOR_MMOTOR_D_MAPPL : LREAL;
	INUMOFCUTLENGTH_LOCK : INT;
	INUMOFCUTLENGTH_INT : INT;
	LRREGPOS_ENDCUT : LREAL := 360;
	LRX_STOPCAMEND : LREAL := 360;
	_XTPCONVERTTPENABLE : BOOL;
	_XSTACKENABLE : BOOL;
	_RC_LRUPPERCORRPOS : LREAL;
	_RC_LRLOWERCORRPOS : LREAL;
	_RC_XENABLE : BOOL;
	_RC_XSYNCHRONISED : BOOL;
	_RC_XTEACHMARKWINDOW : BOOL;
	_RC_XMARKWINDOWOPEN : BOOL;
	_RC_XMARKOUTOFWINDOW : BOOL;
	_RC_XMARKNOTDETECTED : BOOL;
	_RC_XMARKWINDOWTEACHED : BOOL;
	_RC_LRAVERAGEGEARFACTORCORR : LREAL;
	_RC_XGEARFACTORCORRLIMITED : BOOL;
	_RC_LRPOSOUT : LREAL;
	_RC_LRACTVEL : LREAL;
	_RC_XERROR : BOOL;
	_RC_WERRORID : WORD;
	_RC_XLIMITACTIVE : BOOL;
	_RC_LRACTMARKERROR : LREAL;
	_RC_LRACTMARKDIST : LREAL;
	_RC_XINITDONE : BOOL;
	_RC_XCORRACTIVE : BOOL;
	_RC_XMARKRECEIVED : BOOL;
	_RC_LRREGMARKPOS : LREAL;
	_LRREGISTERCNTRFACTOR : LREAL;
	_LRREGISTERCNTRDELAYACTSET : LREAL;
	_RC_XSETREGPOS2MASTERPOS : BOOL;
	_LRTPAXISDELAYCYCLE : LREAL;
	_LRTPDELAYCYCLESACTPOS : LREAL;
	_DWTPAXISDELAYCYCLE : DWORD;
	_LRRESIDUAL : LREAL;
	LRACTMARKPOSDIFF : LREAL;
	FM_REGISTERCONTROLSTATE : L_TF1P_RegisterControlState;
	FB_TPCONVERTTP : L_TT1P_CalculateTPOnMaterialPos := STRUCT(xNoMarkStack := TRUE);
	ITPCONVERTTPENABLECNTR : INT;
	FB_SETTORQUE1 : L_MC1P_SetTorqueOffset;
	FB_STACK : L_MB1P_Stack;
	WRESTART_LOCK : WORD;
	SCCAMTABLE_INT : MC_Cam_REF;
	SCSETXPROFILE_TEMP : L_MC2P_AxisProfile;
	SCSETYPROFILE_TEMP : L_MC2P_AxisProfile;
	PCAMDATA : POINTER TO L_MC2P_CamData;
	C_INUMOFCUTLENGTH : INT := 10;
END_VAR
END_FUNCTION_BLOCK

METHOD CALL_ALLOCPOINTADRBASEEXTENSION
END_METHOD

METHOD CALL_ERRORHANDLER
END_METHOD

METHOD CALL_ERRORHANDLER_STATECUTTING
END_METHOD

METHOD CALL_FBMETHODS
END_METHOD

METHOD CALL_FBMETHODS_BEFOREFLEXCAM
END_METHOD

METHOD CALL_FB_SETTORQUE
END_METHOD

METHOD CALL_FB_SETTORQUE_INPUT
END_METHOD

METHOD CALL_FB_STACK
END_METHOD

METHOD CALL_FB_STACK_INPUT
END_METHOD

METHOD CALL_FB_TPCONVERTTP
END_METHOD

METHOD CALL_FB_TPCONVERTTP_INPUT
END_METHOD

METHOD CALL_FM_CAMCREATOR_STANDSTILL
END_METHOD

METHOD CALL_FM_CAMCREATOR_STOP
END_METHOD

METHOD CALL_FM_CAMCREATORS
END_METHOD

METHOD CALL_FM_FLEXCAM
END_METHOD

METHOD CALL_FM_FLEXCAM_INPUT
END_METHOD

METHOD CALL_FM_REGISTERCONTROL
END_METHOD

METHOD CALL_FM_REGISTERCONTROL_INPUT
END_METHOD

METHOD CALL_FUN_GETSCALING
END_METHOD

METHOD CALL_INITDONE
END_METHOD

METHOD CALL_INITROUTINE
END_METHOD

METHOD CALL_INTERNALCTRL
END_METHOD

METHOD CALL_INTERNALCTRLBASEEXTENSION
END_METHOD

METHOD CALL_OUTPUT
END_METHOD

METHOD CALL_OUTPUTMINMAXVALUES
END_METHOD

METHOD CALL_OUTPUT_SF
END_METHOD

METHOD CALL_RESETCOMMANDS
END_METHOD

METHOD CALL_RESETOUTPUT
END_METHOD

METHOD CALL_RESETWARNINGS
END_METHOD

METHOD CALL_TPCOMPENSATION
END_METHOD

METHOD CALL_CALCCAM_RESTARTFROMSTOPCAM
END_METHOD

METHOD CALL_CALCCAM_STANDSTILL
END_METHOD

METHOD CALL_CALCCAM_STOP
END_METHOD

METHOD CALL_CALCSYNCARRAY_AP10STOPCAM
END_METHOD

METHOD CALL_CHECKARRAYOFCUTLENGTHCHANGES
END_METHOD

METHOD CALL_CHECKCUTPRODUCTFORMAT
END_METHOD

METHOD CALL_CHECKCUTTINGPARCHANGES
END_METHOD

METHOD CALL_CHECKRESTARTFROMSTOPCAM
END_METHOD

METHOD CALL_INIT_FLEXCAM
END_METHOD

METHOD CALL_LOCKCAMTABLE
END_METHOD

METHOD CALL_LOCKCROSSCUTTERPAR
END_METHOD

METHOD CALL_LOCKCUTTINGMODE
END_METHOD

METHOD CALL_LOCKCUTTINGPAR
END_METHOD

METHOD CALL_LOCKCUTTINGPAR_ECCMODE_2
END_METHOD

METHOD CALL_LOCKCUTTINGPAR_ECCMODE_3
END_METHOD

METHOD CALL_LOCKREGISTERCONTROLPAR
END_METHOD

METHOD CALL_PREAPAREARRAYOFCUTLENGTH
END_METHOD

METHOD CALL_PREPARENEXTCUT_ECCMODEPAR
END_METHOD

METHOD CALL_PREPARENEXTCUT_ECCMODEPAR_ECCMODE_2
END_METHOD

METHOD CALL_PREPARENEXTCUT_ECCMODEPAR_ECCMODE_3
END_METHOD

METHOD CALL_CP_000_CYCLIC
END_METHOD

METHOD CALL_CP_001_INIT
END_METHOD

METHOD CALL_CP_144_EXIT_SYNC_PHASE
END_METHOD

METHOD CALL_CP_148_HOLD_IN_PARK_POS
END_METHOD

METHOD CALL_CP_148_HOLD_IN_PARK_POS_CONTINUECUTTING
END_METHOD

METHOD CALL_CP_148_HOLD_IN_PARK_POS_ENDOFPROFILE
END_METHOD

METHOD CALL_CP_801_WAIT_OF_NEXT_CUT
END_METHOD

METHOD CALL_CP_802_STOP_IN_PARK_POS
END_METHOD

METHOD CALL_CP_900_DONE
END_METHOD

METHOD CALL_CUTTING_PROCESS
END_METHOD

METHOD CALL_S000_CYCLIC
END_METHOD

METHOD CALL_S002_READY
END_METHOD

METHOD CALL_S030_SYNCHRONISING_POS
END_METHOD

METHOD CALL_S030_SYNCHRONISING_POS_ECCMODESELECT
END_METHOD

METHOD CALL_S030_SYNCHRONISING_POS_ECCMODE_2
END_METHOD

METHOD CALL_S032_POSITIONING_TO_START_POS
END_METHOD

METHOD CALL_S999_ERROR
END_METHOD

(* ---- _TM_ELECTRICALSHAFTPOSBASE.fb ---- *)
FUNCTION_BLOCK _TM_ELECTRICALSHAFTPOSBASE EXTENDS _TM_MotionControl
VAR_OUTPUT
	PPAR : POINTER TO _scPar_TM_ElectricalShaftPosHigh;
	PSF : POINTER TO _scSF_TM_ElectricalShaftPosHigh;
	PAP : POINTER TO _scAP_TM_ElectricalShaftPosHigh;
END_VAR
VAR_IN_OUT
	MASTERAXIS : AXIS_REF;
	SLAVEAXIS : AXIS_REF;
	XSYNCPOS : BOOL;
	LRSETOFFSETSLAVE : LREAL;
	LRACTVEL : LREAL;
	LRACTPOS : LREAL;
	LROFFSET : LREAL;
END_VAR
VAR
	SCPAR_INT : _scPar_TM_ElectricalShaftPosHigh;
	XSYNCPOS_INT : BOOL;
	LRSETOFFSETSLAVE_INT : LREAL;
	LROFFSET_STORE : LREAL;
	_XSYNCDRIVEENABLE : BOOL;
	_XSYNCDRIVESYNCPOS : BOOL;
	_LRSNYCDRIVESETSLAVEPOSOUT : LREAL;
	_LRSYNCDRIVESETOFFSET : LREAL;
	_LRSYNCDRIVESETOFFSETOUT : LREAL;
	_XLOADSTARTSLAVEPOS : BOOL;
	_LRSTARTSLAVEPOS : LREAL;
	_XLOADGEARBOXPOS : BOOL;
	_LRLOADGEARBOXPOS : LREAL;
	_XLOADOFFSETSYNC : BOOL;
	_LRLOADOFFSETSYNC : LREAL;
	MP03_LRSETGEARBOXPOSOUT : LREAL;
	FM_SYNCHRONIZEDDRIVEBASE1 : L_TF1P_SyncDrivePosBase;
	FB_AXISCONTROLBYPOS : L_MC1P_ControlSetValues;
END_VAR
END_FUNCTION_BLOCK

METHOD CALL_FM_SYNCHRONIZEDDRIVE
END_METHOD

METHOD CALL_FM_SYNCHRONIZEDDRIVE_INPUT
END_METHOD

METHOD CALL_ABC
END_METHOD

METHOD CALL_ALLOCPOINTADR
END_METHOD

METHOD CALL_AXISCONTROLBYPOS
END_METHOD

METHOD CALL_AXISCONTROLBYPOS_INPUT
END_METHOD

METHOD CALL_CTRLREQACTIVE : BOOL
END_METHOD

METHOD CALL_ERRORHANDLER
END_METHOD

METHOD CALL_FBMETHODS
END_METHOD

METHOD CALL_INITDONE
END_METHOD

METHOD CALL_INITROUTINE
END_METHOD

METHOD CALL_INIT_FM
END_METHOD

METHOD CALL_INTERNALCTRL
END_METHOD

METHOD CALL_OUTPUT
END_METHOD

METHOD CALL_OUTPUT_SF
END_METHOD

METHOD CALL_REQUESTS_EXT
END_METHOD

METHOD CALL_RESETCOMMANDS
END_METHOD

METHOD CALL_RESETOUTPUT
END_METHOD

METHOD CALL_STATEMACHINE
END_METHOD

METHOD CALL_S000_CYCLIC
END_METHOD

METHOD CALL_S002_READY
END_METHOD

METHOD CALL_S030_SYNCHRONISING_POS
END_METHOD

METHOD CALL_S031_POS_IS_SYNCHRONISED
END_METHOD

METHOD CALL_S996_STOP
END_METHOD

METHOD CALL_S999_ERROR
END_METHOD

METHOD CALL_T002_READY
END_METHOD

METHOD CALL_T030_SYNCHRONISING_POS
END_METHOD

METHOD CALL_T031_POS_IS_SYNCHRONISED
END_METHOD

(* ---- _TM_ELECTRICALSHAFTPOSHIGH.fb ---- *)
FUNCTION_BLOCK _TM_ELECTRICALSHAFTPOSHIGH EXTENDS _TM_ElectricalShaftPosState
VAR_IN_OUT
	XSYNCINSTANT : BOOL;
	XSYNCOUTINSTANT : BOOL;
	XSYNCPOSRESTORE : BOOL;
	LRSETOFFSETMASTER : LREAL;
	LROFFSETSYNCPOS : LREAL;
	LROFFSETMASTER : LREAL;
END_VAR
VAR
	_XLOADOFFSET : BOOL;
	XSYNCINSTANT_INT : BOOL;
	XSYNCOUTINSTANT_INT : BOOL;
	XSYNCPOSRESTORE_INT : BOOL;
	_XLOADOFFSETMASTER : BOOL;
	LROFFSETMASTER_STORE : LREAL;
	LRFACTORMASTERTOSLAVE : LREAL;
	_LRSYNCDRIVESETOFFSETOUTMASTER : LREAL;
	_LRSYNCDRIVESETOFFSETMASTER : LREAL;
	LRSETOFFSETMASTER_INT : LREAL;
	FM_SYNCHRONIZEDDRIVEHIGH1 : L_TF1P_SyncDriveRegCtrl;
END_VAR
END_FUNCTION_BLOCK

METHOD CALL_FM_SYNCHRONIZEDDRIVE
END_METHOD

METHOD CALL_FM_SYNCHRONIZEDDRIVE_INPUT
END_METHOD

METHOD CALL_CALCFACTORMASTERTOSLAVE
END_METHOD

METHOD CALL_ERRORHANDLER
END_METHOD

METHOD CALL_INITDONE
END_METHOD

METHOD CALL_INITROUTINE
END_METHOD

METHOD CALL_INIT_FM
END_METHOD

METHOD CALL_INTERNALCTRL
END_METHOD

METHOD CALL_OUTPUT
END_METHOD

METHOD CALL_OUTPUT_SF
END_METHOD

METHOD CALL_REQUESTS_EXT
END_METHOD

METHOD CALL_RESETOUTPUT
END_METHOD

METHOD CALL_S000_CYCLIC
END_METHOD

METHOD CALL_S002_READY
END_METHOD

METHOD CALL_S031_POS_IS_SYNCHRONISED
END_METHOD

METHOD CALL_S036_TRIM_POS_PLUS
END_METHOD

METHOD CALL_S037_TRIM_POS_MINUS
END_METHOD

METHOD CALL_T002_READY
END_METHOD

METHOD CALL_T030_SYNCHRONISING_POS
END_METHOD

METHOD CALL_T031_POS_IS_SYNCHRONISED
END_METHOD

(* ---- _TM_ELECTRICALSHAFTPOSSTATE.fb ---- *)
FUNCTION_BLOCK _TM_ELECTRICALSHAFTPOSSTATE EXTENDS _TM_ElectricalShaftPosBase
VAR_IN_OUT
	XTRIMPOS : BOOL;
	XTRIMNEG : BOOL;
	LROFFSETTRIM : LREAL;
	LROFFSETTOTAL : LREAL;
	XSYNCHRONISED : BOOL;
	XACCDECSYNC : BOOL;
END_VAR
VAR
	XTRIMPOS_INT : BOOL;
	XTRIMNEG_INT : BOOL;
	LROFFSETTRIM_STORE : LREAL;
	_XLOADTRIMOFFSET : BOOL;
	_LRLOADTRIMOFFSET : LREAL;
	_LRSETTRIMOFFSETOUT : LREAL;
	_LRSETTOTALOFFSETOUT : LREAL;
	_XSYNCDRIVESYNCOUTINSTANT : BOOL;
	_XSYNCDRIVETRIMPOS : BOOL;
	_XSYNCDRIVETRIMNEG : BOOL;
	_XSYNCDRIVESYNCOUTDONE : BOOL;
	_LRSYNCDRIVEOFFSETSYNCPOS : LREAL;
	_XSYNCDRIVESYNCHRONISED : BOOL;
	_XSYNCDRIVETRIMBUSY : BOOL;
	_XSYNCDRIVEACCDECSYNC : BOOL;
	MP04_LRSETCLUTCHPOS : LREAL;
	FM_SYNCHRONIZEDDRIVESTATE1 : L_TF1P_SyncDrivePosState;
END_VAR
END_FUNCTION_BLOCK

METHOD CALL_FM_SYNCHRONIZEDDRIVE
END_METHOD

METHOD CALL_FM_SYNCHRONIZEDDRIVE_INPUT
END_METHOD

METHOD CALL_ERRORHANDLER
END_METHOD

METHOD CALL_INITDONE
END_METHOD

METHOD CALL_INITROUTINE
END_METHOD

METHOD CALL_INIT_FM
END_METHOD

METHOD CALL_INTERNALCTRL
END_METHOD

METHOD CALL_OUTPUT
END_METHOD

METHOD CALL_OUTPUT_SF
END_METHOD

METHOD CALL_REQUESTS_EXT
END_METHOD

METHOD CALL_RESETCOMMANDS
END_METHOD

METHOD CALL_RESETOUTPUT
END_METHOD

METHOD CALL_STATEMACHINE
END_METHOD

METHOD CALL_S000_CYCLIC
END_METHOD

METHOD CALL_S030_SYNCHRONISING_POS
END_METHOD

METHOD CALL_S031_POS_IS_SYNCHRONISED
END_METHOD

METHOD CALL_S036_TRIM_POS_PLUS
END_METHOD

METHOD CALL_S037_TRIM_POS_MINUS
END_METHOD

METHOD CALL_T030_SYNCHRONISING_POS
END_METHOD

METHOD CALL_T031_POS_IS_SYNCHRONISED
END_METHOD

(* ---- _TM_ELECTRICALSHAFTVELBASE.fb ---- *)
FUNCTION_BLOCK _TM_ELECTRICALSHAFTVELBASE EXTENDS _TM_MotionControl
VAR_OUTPUT
	PPAR : POINTER TO _scPar_TM_ElectricalShaftVelHigh;
	PSF : POINTER TO _scSF_TM_ElectricalShaftVelHigh;
	PAP : POINTER TO _scAP_TM_ElectricalShaftVelHigh;
END_VAR
VAR_IN_OUT
	MASTERAXIS : AXIS_REF;
	SLAVEAXIS : AXIS_REF;
	XSYNCVEL : BOOL;
	LRSETOFFSET : LREAL;
	LRACTVEL : LREAL;
	LRACTPOS : LREAL;
	LROFFSET : LREAL;
END_VAR
VAR
	SCPAR_INT : _scPar_TM_ElectricalShaftVelHigh;
	XSYNCVEL_INT : BOOL;
	LRSETOFFSET_INT : LREAL;
	LRCOUPLINGX_INT : LREAL;
	DWMODE_INT : DWORD;
	LRCOUPLINGY_INT : LREAL;
	XERROR_MODULOAXISISREQUIRED : BOOL;
	XERROR_INVALIDCOUPLINGMODE : BOOL;
	ETMSTATE_INT_TEMP : L_TT1P_States;
	_XSYNCDRIVEENABLE : BOOL;
	_LRSYNCDRIVESETSLAVEVELOUT : LREAL;
	_LROFFSET : LREAL;
	FM_SYNCHRONIZEDDRIVEBASE1 : L_TF1P_SyncDriveVelBase;
	FB_CONTROLAXISBYVEL : L_MC1P_ControlSetValues := STRUCT(xIgnoreAccForPosCalc := TRUE);
	LRMASTERSETPOSITIONFORSYNC_OLD : LREAL;
END_VAR
END_FUNCTION_BLOCK

METHOD CALL_ALLOCPOINTADR
END_METHOD

METHOD CALL_CTRLREQACTIVE : BOOL
END_METHOD

METHOD CALL_ERRORHANDLER
END_METHOD

METHOD CALL_FBMETHODS
END_METHOD

METHOD CALL_FB_CONTROLAXISBYVEL
END_METHOD

METHOD CALL_FB_CONTROLAXISBYVEL_INPUT
END_METHOD

METHOD CALL_FM_SYNCHRONIZEDDRIVE
END_METHOD

METHOD CALL_FM_SYNCHRONIZEDDRIVE_INPUT
END_METHOD

METHOD CALL_FM_SYNCHRONIZEDDRIVE_RESETFM
END_METHOD

METHOD CALL_INITDONE
END_METHOD

METHOD CALL_INITROUTINE
END_METHOD

METHOD CALL_INTERNALCTRL
END_METHOD

METHOD CALL_OUTPUT
END_METHOD

METHOD CALL_OUTPUT_FM_SYNCHRONIZEDDRIVE
END_METHOD

METHOD CALL_OUTPUT_SF
END_METHOD

METHOD CALL_REQUESTS_EXT
END_METHOD

METHOD CALL_RESETCOMMANDS
END_METHOD

METHOD CALL_RESETOUTPUT
END_METHOD

METHOD CALL_STATEMACHINE
END_METHOD

METHOD CALL_ABC
END_METHOD

METHOD CALL_S002_READY
END_METHOD

METHOD CALL_S041_VEL_IS_SYNCHRONISED
END_METHOD

METHOD CALL_S052_ACC_DEC
END_METHOD

METHOD CALL_S999_ERROR
END_METHOD

METHOD CALL_T002_READY
END_METHOD

METHOD CALL_T041_VEL_IS_SYNCHRONISED
END_METHOD

METHOD CALL_T052_ACC_DEC
END_METHOD

(* ---- _TM_ELECTRICALSHAFTVELHIGH.fb ---- *)
FUNCTION_BLOCK _TM_ELECTRICALSHAFTVELHIGH EXTENDS _TM_ElectricalShaftVelState
VAR_INPUT
	LRSETGROUNDVEL : LREAL := 0;
END_VAR
VAR
	LRSETGROUNDVEL_INT : LREAL := 0.0;
	LRSETGROUNDVEL_OLD : LREAL;
	XVELSYNCOUTTOGROUNDSPEEDBUSY : BOOL;
	_LRSETGROUNDVEL : LREAL;
	XFM_SD_OFFSETBUSY : BOOL;
	_XSYNCHRONISEDGROUNDVEL : BOOL;
	XFM_SD_ACCDECGROUNDVEL : BOOL;
	FM_SYNCHRONIZEDDRIVEHIGH1 : L_TF1P_SyncDriveVelHigh;
END_VAR
END_FUNCTION_BLOCK

METHOD CALL_ERRORHANDLER
END_METHOD

METHOD CALL_FM_SYNCHRONIZEDDRIVE
END_METHOD

METHOD CALL_FM_SYNCHRONIZEDDRIVE_INPUT
END_METHOD

METHOD CALL_FM_SYNCHRONIZEDDRIVE_RESETFM
END_METHOD

METHOD CALL_INTERNALCTRL
END_METHOD

METHOD CALL_OUTPUT
END_METHOD

METHOD CALL_OUTPUT_FM_SYNCHRONIZEDDRIVE
END_METHOD

METHOD CALL_OUTPUT_SF
END_METHOD

METHOD CALL_REQUESTS_EXT
END_METHOD

METHOD CALL_RESETCOMMANDS
END_METHOD

METHOD CALL_RESETOUTPUT
END_METHOD

METHOD CALL_STATEMACHINE
END_METHOD

METHOD CALL_S002_READY
END_METHOD

METHOD CALL_S041_VEL_IS_SYNCHRONISED
END_METHOD

METHOD CALL_S051_GROUNDSPEED
END_METHOD

METHOD CALL_S052_ACC_DEC
END_METHOD

METHOD CALL_T002_READY
END_METHOD

METHOD CALL_T041_VEL_IS_SYNCHRONISED
END_METHOD

METHOD CALL_T051_GROUNDSPEED
END_METHOD

METHOD CALL_T052_ACC_DEC
END_METHOD

(* ---- _TM_ELECTRICALSHAFTVELSTATE.fb ---- *)
FUNCTION_BLOCK _TM_ELECTRICALSHAFTVELSTATE EXTENDS _TM_ElectricalShaftVelBase
VAR_IN_OUT
	XTRIMPOS : BOOL;
	XTRIMNEG : BOOL;
	LROFFSETTRIM : LREAL;
	LROFFSETTOTAL : LREAL;
	XSYNCHRONISED : BOOL;
	XACCDECSYNC : BOOL;
END_VAR
VAR
	XTRIMPOS_INT : BOOL;
	XTRIMNEG_INT : BOOL;
	XTRIMPOS_INT_OLD : BOOL;
	XTRIMNEG_INT_OLD : BOOL;
	_XSYNCVEL : BOOL;
	_XTRIMPOS : BOOL;
	_XTRIMNEG : BOOL;
	_LROFFSETTRIM : LREAL;
	_LROFFSETTOTAL : LREAL;
	_XSYNCOUTDONE : BOOL;
	_XSYNCHRONISED : BOOL;
	_XACCDECSYNC : BOOL;
	_XTRIMBUSY : BOOL;
	FM_SYNCHRONIZEDDRIVESTATE1 : L_TF1P_SyncDriveVelState;
	LRCOUPLINGXOLD : LREAL;
	LRCOUPLINGYOLD : LREAL;
END_VAR
END_FUNCTION_BLOCK

METHOD CALL_ERRORHANDLER
END_METHOD

METHOD CALL_FM_SYNCHRONIZEDDRIVE
END_METHOD

METHOD CALL_FM_SYNCHRONIZEDDRIVE_INPUT
END_METHOD

METHOD CALL_FM_SYNCHRONIZEDDRIVE_RESETFM
END_METHOD

METHOD CALL_INTERNALCTRL
END_METHOD

METHOD CALL_OUTPUT
END_METHOD

METHOD CALL_OUTPUT_SF
END_METHOD

METHOD CALL_RESETCOMMANDS
END_METHOD

METHOD CALL_RESETOUTPUT
END_METHOD

METHOD CALL_STATEMACHINE
END_METHOD

METHOD CALL_S002_READY
END_METHOD

METHOD CALL_S036_TRIM_POS_PLUS
END_METHOD

METHOD CALL_S037_TRIM_POS_MINUS
END_METHOD

METHOD CALL_S041_VEL_IS_SYNCHRONISED
END_METHOD

METHOD CALL_S052_ACC_DEC
END_METHOD

METHOD CALL_S996_STOP
END_METHOD

METHOD CALL_T002_READY
END_METHOD

METHOD CALL_T041_VEL_IS_SYNCHRONISED
END_METHOD

METHOD CALL_T052_ACC_DEC
END_METHOD

(* ---- _TM_FLEXCAMBASE.fb ---- *)
FUNCTION_BLOCK _TM_FLEXCAMBASE EXTENDS _TM_MotionControl
VAR_OUTPUT
	PAP : POINTER TO _scAP_TM_FlexCamHigh;
	PPAR : POINTER TO _scPar_TM_FlexCamHigh;
	PSF : POINTER TO _scSF_TM_FlexCamHigh;
END_VAR
VAR_IN_OUT
	MASTERAXIS : AXIS_REF;
	SLAVEAXIS : AXIS_REF;
	XENABLEHWLIMIT : BOOL;
	XHWLIMITPOS : BOOL;
	XHWLIMITNEG : BOOL;
	XSYNCCAM : BOOL;
	XSYNCOUTINSTANT : BOOL;
	XCAMCHANGEINSTANT : BOOL;
	LRSETOFFSETMASTER : LREAL;
	LRSETOFFSETSLAVE : LREAL;
	LRSETSCALINGMASTER : LREAL;
	LRSETSCALINGSLAVE : LREAL;
	CAMTABLE1 : MC_CAM_REF;
	XHWLIMITSWITCHNEG : BOOL;
	XHWLIMITSWITCHPOS : BOOL;
	XSWLIMITENABLED : BOOL;
	XSWLIMITSWITCHACTIVE : BOOL;
	XCAMSYNCHRONISED : BOOL;
	XACCDECSYNC : BOOL;
	XENDOFPROFILE : BOOL;
	LRSETXPOSOUT : LREAL;
	LRSETXVELOUT : LREAL;
	LRSETXACCOUT : LREAL;
	LRSETYPOSOUT : LREAL;
	LRSETYVELOUT : LREAL;
	LRSETYACCOUT : LREAL;
	LRACTSLAVEPOS : LREAL;
	LRACTSLAVEVEL : LREAL;
	LRSETOFFSETMASTEROUT : LREAL;
	LRSETOFFSETSLAVEOUT : LREAL;
	LRSLAVEMAXPOS : LREAL;
	LRSLAVEMINPOS : LREAL;
	LRSLAVEMAXVEL : LREAL;
	LRSLAVEMAXACC : LREAL;
END_VAR
VAR
	XSYNCCAM_INT : BOOL;
	XSYNCOUTINSTANT_INT : BOOL;
	XCAMCHANGEINSTANT_INT : BOOL;
	LRSETOFFSETMASTER_INT : LREAL;
	LRSETOFFSETSLAVE_INT : LREAL;
	LRSETSCALINGMASTER_INT : LREAL;
	LRSETSCALINGSLAVE_INT : LREAL;
	SCPAR_INT : _scPar_TM_FlexCamHigh;
	XENABLEHWLIMIT_INT : BOOL;
	XHWLIMITPOS_INT : BOOL;
	XHWLIMITNEG_INT : BOOL;
	XHOMEEXECUTE_OLD : BOOL;
	XCAMCHANGEINSTANT_OLD : BOOL;
	LRMASTERVEL_OLD : LREAL;
	LRMASTERVEL_OLD2 : LREAL;
	LRMASTERPOS_OLD : LREAL;
	XMASTERAXISENABLED : BOOL;
	XMASTERAXISENABLED_OLD : BOOL;
	XMASTERIS_FREEENCODER : BOOL;
	XINVALIDMASTER : BOOL := FALSE;
	XCRITICALERROR : BOOL;
	XCOMMUNICATION : BOOL;
	CAMTABLE_INIT : MC_CAM_REF;
	XVISHOMEPARACTIVE : BOOL;
	XCAMTABLEINTERNALVALID : BOOL;
	CAMTABLEINTERNAL : MC_CAM_REF;
	PCAMDATA : POINTER TO L_MC2P_CamData;
	_XFC_ENABLE : BOOL;
	_LRFC_SETXPOSOUT : LREAL;
	_LRFC_SETXVELOUT : LREAL;
	_LRFC_SETXACCOUT : LREAL;
	_LRFC_SETYPOSOUT : LREAL;
	_LRFC_SETYVELOUT : LREAL;
	_LRFC_SETYACCOUT : LREAL;
	_LRFC_SETOFFSETMASTEROUT : LREAL;
	_LRFC_SETOFFSETSLAVEOUT : LREAL;
	_XFC_CRITICALCYCLE : BOOL;
	_XFC_ENDOFPROFILE : BOOL;
	_XFC_ACCDECSYNC : BOOL;
	_XFC_CAMSYNCHRONISED : BOOL;
	_XFC_BUSY : BOOL;
	_XFC_DONE : BOOL;
	_LRFC_SETSLAVEPOSOUT : LREAL;
	_LRFC_SETSLAVEVELOUT : LREAL;
	_LRFC_SETSLAVEACCOUT : LREAL;
	LRENDOFPROFILEWINDOWSIZE : LREAL := 0;
	MP03_LRCONVERTMASTERTOXPOS : LREAL;
	MP04_LRCAMPROFILERPOSOUT : LREAL;
	MP05_LRSETYPOS : LREAL;
	MP06_LRCONVERTYTOSLAVEPOS : LREAL;
	MP00_LWENDOFPROFILECHECKSUM : LWORD;
	MP07_XENDOFPROFPOSITIVE : BOOL;
	MP08_XENDOFPROFNEGATIVE : BOOL;
	SCSETXPROFILE : L_MC2P_AxisProfile;
	SCSETYPROFILE : L_MC2P_AxisProfile;
	FB_CAMBASIC : L_MC2P_CamBasic;
	FB_CONTROLSETVALUES : L_MC1P_ControlSetValues;
	FB_CAMTABLEINFO1 : L_MB1P_CamTableInfo;
	FB_HWLIMITAXIS : L_MC1P_HWLimitSwitchInterface;
END_VAR
END_FUNCTION_BLOCK

METHOD CALL_ALLOCPOINTADR
END_METHOD

METHOD CALL_AXISCONTROLBYPOS
END_METHOD

METHOD CALL_AXISCONTROLBYPOS_INPUT
END_METHOD

METHOD CALL_CAMBOUNDS
END_METHOD

METHOD CALL_CTRLREQACTIVE : BOOL
END_METHOD

METHOD CALL_CURVESKETCHING
END_METHOD

METHOD CALL_ERRORHANDLER
END_METHOD

METHOD CALL_FBMETHODS
END_METHOD

METHOD CALL_FB_CAMBASIC
END_METHOD

METHOD CALL_FB_HWLIMITAXIS
END_METHOD

METHOD CALL_FM_CAMTABLEINFO1
END_METHOD

METHOD CALL_FM_FLEXCAM
END_METHOD

METHOD CALL_FM_FLEXCAM_INPUT
END_METHOD

METHOD CALL_FIRSTCYCLE
END_METHOD

METHOD CALL_INITDONE
END_METHOD

METHOD CALL_INITROUTINE
END_METHOD

METHOD CALL_INTERNALCTRL
END_METHOD

METHOD CALL_LIMITEDINPUT
END_METHOD

METHOD CALL_OUTPUT
END_METHOD

METHOD CALL_OUTPUTMINMAXVALUES
END_METHOD

METHOD CALL_OUTPUTMINMAXVALUESMODULOOVERRUN
END_METHOD

METHOD CALL_OUTPUTMINMAXVALUESOFCAMTABLES1
END_METHOD

METHOD CALL_OUTPUT_SF
END_METHOD

METHOD CALL_REQUESTS_EXT
END_METHOD

METHOD CALL_RESETCOMMANDS
END_METHOD

METHOD CALL_RESETOUTPUT
END_METHOD

METHOD CALL_STATEMACHINE
END_METHOD

METHOD CALL_ABC
END_METHOD

METHOD CAMREFCHANGED : BOOL
VAR_IN_OUT
	CAMREFNEW : MC_CAM_REF;
	CAMREFOLD : MC_CAM_REF;
END_VAR
END_METHOD

METHOD CAMREFVALID : BOOL
VAR_INPUT
	CAMREF : MC_CAM_REF;
END_VAR
END_METHOD

METHOD GET_INTERNCAMTABLE : MC_CAM_REF
END_METHOD

METHOD GET_ECAMTYPE : L_MC2P_CamType
END_METHOD

METHOD GET_LRCAMXEND : LREAL
END_METHOD

METHOD GET_LRCAMXSTART : LREAL
END_METHOD

METHOD GET_LRCAMYEND : LREAL
END_METHOD

METHOD GET_LRCAMYSTART : LREAL
END_METHOD

METHOD GET_XCOMMUNICATION : BOOL
END_METHOD

METHOD RESET_SYSTEMFAULT
END_METHOD

METHOD SET_SYSTEMFAULT
VAR_INPUT
	IN : L_IE1P_Error;
END_VAR
END_METHOD

METHOD SET_ESTATE
VAR_INPUT
	IN : L_TT1P_States;
END_VAR
END_METHOD

METHOD CALL_S000_CYCLIC
END_METHOD

METHOD CALL_S002_READY
END_METHOD

METHOD CALL_S112_CAMMING
END_METHOD

METHOD CALL_S996_STOP
END_METHOD

METHOD CALL_S999_ERROR
END_METHOD

METHOD CALL_T002_READY
END_METHOD

(* ---- _TM_FLEXCAMBASEEXTENSION.fb ---- *)
FUNCTION_BLOCK _TM_FLEXCAMBASEEXTENSION EXTENDS _TM_FlexCamBase
VAR
	FM_FLEXCAMBASE1 : L_MC2P_FlexCamBase;
END_VAR
END_FUNCTION_BLOCK

METHOD CALL_ERRORHANDLER
END_METHOD

METHOD CALL_FM_FLEXCAM
END_METHOD

METHOD CALL_FM_FLEXCAM_INPUT
END_METHOD

METHOD CALL_OUTPUTMINMAXVALUES
END_METHOD

METHOD CALL_OUTPUTMINMAXVALUESOFCAMTABLES1
END_METHOD

METHOD GET_INTERNCAMTABLE : MC_CAM_REF
END_METHOD

METHOD GET_LRCAMXEND : LREAL
END_METHOD

METHOD GET_LRCAMXSTART : LREAL
END_METHOD

METHOD GET_LRCAMYEND : LREAL
END_METHOD

METHOD GET_LRCAMYSTART : LREAL
END_METHOD

(* ---- _TM_FLEXCAMSTATE.fb ---- *)
FUNCTION_BLOCK _TM_FLEXCAMSTATE EXTENDS _TM_FlexCamBase
VAR_OUTPUT
	ESETCAMTABLEOUT : L_TT1P_CamTable;
END_VAR
VAR_IN_OUT
	CAMTABLE2 : MC_CAM_REF;
	CAMTABLE3 : MC_CAM_REF;
	CAMTABLE4 : MC_CAM_REF;
	ESETCAMTABLE : L_TT1P_CamTable;
	XCAMSEQUENCER : BOOL;
	XCAMSEQUENCERACTIVE : BOOL;
END_VAR
VAR
	ESETCAMTABLE_INT : L_TT1P_CamTable;
	XCAMSEQUENCER_INT : BOOL;
	XSLAVEABSOLUTE_OLD : BOOL;
	XUPDATECURVE : BOOL;
	_XMCS_ENABLE : BOOL;
	_MCS_CAMTABLEOUT : MC_CAM_REF;
	FM_FLEXCAMSTATE1 : L_MC2P_FlexCamState;
	FB_MULTICAMSEQUENCER1 : L_MB1P_MultiCamSequencer;
	FB_CAMTABLEINFO2 : L_MB1P_CamTableInfo;
	FB_CAMTABLEINFO3 : L_MB1P_CamTableInfo;
	FB_CAMTABLEINFO4 : L_MB1P_CamTableInfo;
END_VAR
END_FUNCTION_BLOCK

METHOD CALL_CURVESKETCHING
END_METHOD

METHOD CALL_ERRORHANDLER
END_METHOD

METHOD CALL_FBMETHODS
END_METHOD

METHOD CALL_FM_CAMTABLEINFO2
END_METHOD

METHOD CALL_FM_CAMTABLEINFO3
END_METHOD

METHOD CALL_FM_CAMTABLEINFO4
END_METHOD

METHOD CALL_FM_FLEXCAM
END_METHOD

METHOD CALL_FM_FLEXCAM_INPUT
END_METHOD

METHOD CALL_FM_MULTICAMSEQUENCER
END_METHOD

METHOD CALL_FM_MULTICAMSEQUENCER_INPUT
END_METHOD

METHOD CALL_FIRSTCYCLE
END_METHOD

METHOD CALL_INTERNALCTRL
END_METHOD

METHOD CALL_OUTPUT
END_METHOD

METHOD CALL_OUTPUTMINMAXVALUES
END_METHOD

METHOD CALL_OUTPUTMINMAXVALUESOFCAMTABLES1
END_METHOD

METHOD CALL_OUTPUTMINMAXVALUESOFCAMTABLES1_2_3_4
END_METHOD

METHOD CALL_OUTPUT_SF
END_METHOD

METHOD CALL_RESETCOMMANDS
END_METHOD

METHOD CALL_RESETCOMMANDSFLEXCAM
END_METHOD

METHOD CALL_RESETOUTPUT
END_METHOD

METHOD GET_INTERNCAMTABLE : MC_CAM_REF
END_METHOD

METHOD GET_LRCAMXEND : LREAL
END_METHOD

METHOD GET_LRCAMXSTART : LREAL
END_METHOD

METHOD GET_LRCAMYEND : LREAL
END_METHOD

METHOD GET_LRCAMYSTART : LREAL
END_METHOD

(* ---- _TM_FLYINGSAWBASE.fb ---- *)
FUNCTION_BLOCK _TM_FLYINGSAWBASE EXTENDS _TM_MotionControl
VAR_OUTPUT
	PPAR : POINTER TO _scPar_TM_FlyingSawHigh;
	PSF : POINTER TO _scSF_TM_FlyingSawHigh;
	PAP : POINTER TO _scAP_TM_FlyingSawHigh;
END_VAR
VAR_IN_OUT
	MASTERAXIS : AXIS_REF;
	SLAVEAXIS : AXIS_REF;
	XENABLEHWLIMIT : BOOL;
	XHWLIMITPOS : BOOL;
	XHWLIMITNEG : BOOL;
	XSTARTFLYINGSAW : BOOL;
	XSYNCININSTANT : BOOL;
	XEXECUTENEXTCUT : BOOL;
	XEXECUTEGAP : BOOL;
	LRCUTTINGLENGTH : LREAL;
	XSETMATERIALCOUNTER : BOOL;
	XHWLIMITSWITCHNEG : BOOL;
	XHWLIMITSWITCHPOS : BOOL;
	XSWLIMITENABLED : BOOL;
	XSWLIMITSWITCHACTIVE : BOOL;
	XSYNCHRONIZED : BOOL;
	XACCDECSYNC : BOOL;
	XPOSITIONING : BOOL;
	XINPOSITION : BOOL;
	LRACTPOS : LREAL;
	LRACTVEL : LREAL;
	LRACTFOLLOWINGERROR : LREAL;
	LRMATERIALCOUNTER : LREAL;
	LRTARGETPOS : LREAL;
	LRCUTGAP : LREAL;
END_VAR
VAR
	SCPAR_INT : _scPar_TM_FlyingSawHigh;
	XSTARTFLYINGSAW_INT : BOOL;
	XSYNCININSTANT_INT : BOOL;
	LRSETOFFSETSLAVE_INT : LREAL;
	XSETMATERIALCOUNTER_INT : BOOL;
	XEXECUTENEXTCUT_INT : BOOL;
	XENABLEHWLIMIT_INT : BOOL;
	XHWLIMITPOS_INT : BOOL;
	XHWLIMITNEG_INT : BOOL;
	XEXECUTEGAP_INT : BOOL;
	LROFFSET_STORE : LREAL;
	FB_MATERIALCOUNTER : L_MB1P_MaterialCounter;
	FB_CALCULATETARGETPOS : L_TT1P_CalculateTargetPos;
	FB_PROCESSCONTROL : L_TT1P_ProcessControl;
	FB_POSPROFILERCLUTCH : L_MB1P_PosProfilerClutchState;
	FB_POSPROFILER_INIT : L_MC1P_PosProfiler;
	SCPROFILEPARAMETER : L_MC1P_ProfileParameter;
	FB_CONTROLSETVALUES : L_MC1P_ControlSetValues;
	FB_HWLIMITAXIS : L_MC1P_HWLimitSwitchInterface;
	WSTEPPER : WORD;
	LRSTARTPOSOUT : LREAL;
	LRSTARTPOSOUT2 : LREAL;
	LRACCDIST : LREAL;
	LRACCTIME : LREAL;
	XERRORSTOP : BOOL;
	LRDECDIST : LREAL;
	LRDECTIME : LREAL;
	LRMASTERPOS1 : LREAL;
	LRMASTERPOS2 : LREAL;
	LRSLAVEPOS1 : LREAL;
	LRSLAVEPOS2 : LREAL;
	XSYNCHRONIZEDOLD : BOOL;
	WSTEPPER1 : WORD;
	LRCUTGAP_INT : LREAL;
	XACCDECSYNC_OLD : BOOL;
	XGAPDONE : BOOL;
	WSTEPPER2 : WORD;
	LRCUTTINGLENGTH_INT : LREAL;
	LRJERK_INT : LREAL;
	LRDIST_INT : LREAL;
	EMODEFLYINGSAW_INT : L_TT1P_eModesFlyingSaw := L_TT1P_eModesFlyingSaw.LengthControlled;
	XRESETMARKSTACK_INT : BOOL;
	XTEST : BOOL;
END_VAR
END_FUNCTION_BLOCK

METHOD CALL_ABC
END_METHOD

METHOD CALL_ALLOCPOINTADR
END_METHOD

METHOD CALL_CALCULATECUTTINGLENGTH
END_METHOD

METHOD CALL_CTRLREQACTIVE : BOOL
END_METHOD

METHOD CALL_ERRORHANDLER
END_METHOD

METHOD CALL_INITDONE
END_METHOD

METHOD CALL_INITROUTINE
END_METHOD

METHOD CALL_INTERNALCTRL
END_METHOD

METHOD CALL_OUTPUT
END_METHOD

METHOD CALL_OUTPUT_SF
END_METHOD

METHOD CALL_REQUESTS_EXT
END_METHOD

METHOD CALL_RESETCOMMANDS
END_METHOD

METHOD CALL_RESETOUTPUT
END_METHOD

METHOD CALL_STATEMACHINE
END_METHOD

METHOD CALL_FBMETHODS
END_METHOD

METHOD CALL_FB_CALCULATETPONMATERIALPOS
END_METHOD

METHOD CALL_FB_CALCULATETPONMATERIALPOSINPUTS
END_METHOD

METHOD CALL_FB_CALCULATETARGETPOS
END_METHOD

METHOD CALL_FB_CALCULATETARGETPOSINPUTS
END_METHOD

METHOD CALL_FB_CONTROLSETVALUESINPUTS
END_METHOD

METHOD CALL_FB_CONTROLSETVALUES
END_METHOD

METHOD CALL_FB_HWLIMITAXISINPUTS
END_METHOD

METHOD CALL_FB_HWLIMITAXIS
END_METHOD

METHOD CALL_FB_INPOSITION
END_METHOD

METHOD CALL_FB_INPOSITIONINPUTS
END_METHOD

METHOD CALL_FB_MATERIALCOUNTERINPUTS
END_METHOD

METHOD CALL_FB_MATERIALCOUNTER
END_METHOD

METHOD CALL_FB_POSPROFILERCLUTCH
END_METHOD

METHOD CALL_FB_POSPROFILERCLUTCHINPUTS
END_METHOD

METHOD CALL_FB_PROCESSCONTROL
END_METHOD

METHOD CALL_FB_PROCESSCONTROLINPUTS
END_METHOD

METHOD CALL_S000_CYCLIC
END_METHOD

METHOD CALL_S002_READY
END_METHOD

METHOD CALL_S030_SAW_IN_PROCESS
END_METHOD

METHOD CALL_S996_STOP
END_METHOD

METHOD CALL_S999_ERROR
END_METHOD

METHOD CALL_T002_READY
END_METHOD

METHOD CALL_T030_SAW_IN_PROCESS
END_METHOD

METHOD CALL_S000_STARTSAW
END_METHOD

METHOD CALL_S020_SAWSYNCHRONIZED
END_METHOD

METHOD CALL_S030_MOVETOLOWERLIMIT
END_METHOD

METHOD CALL_S040_WAITINGFORNEXTCUT
END_METHOD

(* ---- _TM_FLYINGSAWSTATE.fb ---- *)
FUNCTION_BLOCK _TM_FLYINGSAWSTATE EXTENDS _TM_FlyingSawBase
VAR_IN_OUT
	XMOVETOPARKPOS : BOOL;
	XRESUMETARGETPOS : BOOL;
	XRESETMARKSTACK : BOOL;
	XMARKRECEIVE : BOOL;
	LRACTMARKPOSIN : LREAL;
	BYREMAINMARKSTACK : BYTE;
END_VAR
VAR
	FB_CALCULATETPCOMPENSATIONFACTOR : L_MB1P_CalculateTpCompensationFactor;
	FB_CALCULATETPONMATERIALPOS : L_TT1P_CalculateTPOnMaterialPos;
	FB_INPOSITION : L_TT1P_InPosition;
	FB_SR : SR;
	R_TRIG3 : R_TRIG;
	F_TRIG1 : F_TRIG;
	FB_SR2 : SR;
	LRSYNCOUTPOS : LREAL;
	XNEXTCUT_IP : BOOL;
	XMOVETOPARKPOS_INT : BOOL;
	XRESUMETARGETPOS_INT : BOOL;
	WSTEPPERSKPCUT : INT;
	XSYNCINSTANT_IP : BOOL;
	XFIRSTTP : BOOL;
	XMODECHANGE : BOOL;
	XMODECHANGE_OLD : BOOL;
	EMODEFLYINGSAW_OLD : L_TT1P_eModesFlyingSaw;
	PAXISREAL : POINTER TO _AXIS_REF_REAL;
	BYTEST : BYTE;
	LRRANGEOFTOLERANCE : LREAL;
	_LRREGISTERCNTRFACTOR : LREAL;
	_LRTPAXISDELAYCYCLE : LREAL;
	_LRTPDELAYCYCLESACTPOS : LREAL;
	_DWTPAXISDELAYCYCLE : DWORD;
	_LRRESIDUAL : LREAL;
END_VAR
END_FUNCTION_BLOCK

METHOD CALL_ALLOCPOINTADR
END_METHOD

METHOD CALL_ERRORHANDLER
END_METHOD

METHOD CALL_INTERNALCTRL
END_METHOD

METHOD CALL_OUTPUT
END_METHOD

METHOD CALL_OUTPUT_SF
END_METHOD

METHOD CALL_REQUESTS_EXT
END_METHOD

METHOD CALL_STATEMACHINE
END_METHOD

METHOD CALL_TPVALID
END_METHOD

METHOD CALL_FBMETHODS
END_METHOD

METHOD CALL_FB_CALCULATETPONMATERIALPOS
END_METHOD

METHOD CALL_FB_CALCULATETPONMATERIALPOSINPUTS
END_METHOD

METHOD CALL_FB_CALCULATETARGETPOSINPUTS
END_METHOD

METHOD CALL_FB_CALCULATETPCOMPENSATIONFACTOR
END_METHOD

METHOD CALL_FB_INPOSITIONINPUTS
END_METHOD

METHOD CALL_FB_INPOSITION
END_METHOD

METHOD CALL_FB_POSPROFILERCLUTCHINPUTS
END_METHOD

METHOD CALL_FB_PROCESSCONTROLINPUTS
END_METHOD

METHOD CALL_S000_CYCLIC
END_METHOD

METHOD CALL_S002_READY
END_METHOD

METHOD CALL_S003_HOMING
END_METHOD

METHOD CALL_S010_JOGGING
END_METHOD

METHOD CALL_S030_SAW_IN_PROCESS
END_METHOD

METHOD CALL_S040_MOVE_TO_PARKPOS
END_METHOD

METHOD CALL_S996_STOP
END_METHOD

METHOD CALL_T002_READY
END_METHOD

METHOD CALL_T030_SAW_IN_PROCESS
END_METHOD

METHOD CALL_S000_STARTSAW
END_METHOD

METHOD CALL_S040_WAITINGFORNEXTCUT
END_METHOD

(* ---- _TM_MOTIONCONTROL.fb ---- *)
FUNCTION_BLOCK _TM_MOTIONCONTROL EXTENDS _TM_MotionControlBase
VAR_OUTPUT
	EERRORID : L_IE1P_Error;
END_VAR
VAR_IN_OUT
	SCCTRLABC : scCtrl_ABC;
	XRESETERROR : BOOL;
	XREGULATORON : BOOL;
	XSTOP : BOOL;
	XHALT : BOOL;
	SCACCESSPOINTS : _scAP_TM_MotionControl;
	XJOGPOS : BOOL;
	XJOGNEG : BOOL;
	XHOMEEXECUTE : BOOL;
	XHOMEABSSWITCH : BOOL;
	SCPAR : _scPar_TM_MotionControl;
	SCSTATUSABC : scStatus_ABC;
	XERROR : BOOL;
	XWARNING : BOOL;
	SCERRORINFO : L_TT1P_scErrorInfo;
	XAXISENABLED : BOOL;
	SCSIGNALFLOW : _scSF_TM_MotionControl;
	XBUSY : BOOL;
	XDONE : BOOL;
	XISHOMED : BOOL;
END_VAR
VAR
	SCCTRLABC_INT : scCtrl_ABC;
	XJOGPOS_INT : BOOL;
	XJOGNEG_INT : BOOL;
	XHOMEEXECUTE_INT : BOOL;
	XHOMEABSSWITCH_INT : BOOL;
	PPARABC : POINTER TO _scPar_TM_MotionControl;
	PPARJOGGING : POINTER TO _scPar_TM_MotionControlBase;
	PPARHOMING : POINTER TO _scPar_TM_MotionControlState;
	PABCCTRL : POINTER TO scCtrl_ABC;
	XAXISNOTENABLED : BOOL;
	XINVALIDINPUTJOGPOSJOGNEG : BOOL;
	XINTERRUPTHOMINGBYHALT : BOOL;
	ABC : L_MC1P_AxisBasicControl;
END_VAR
END_FUNCTION_BLOCK

METHOD CALL_ABCCTRLREQACTIVE : BOOL
END_METHOD

METHOD CALL_ABCGENERALSETTINGS
END_METHOD

METHOD CALL_ALLOCPOINTADR
END_METHOD

METHOD CALL_ERRORHANDLER
END_METHOD

METHOD CALL_ERRORHANDLER_SCERRORINFO
END_METHOD

METHOD CALL_FBMETHODS
END_METHOD

METHOD CALL_FIRSTCYCLE
END_METHOD

METHOD CALL_INITROUTINE
END_METHOD

METHOD CALL_INTERNALCTRL
END_METHOD

METHOD CALL_OUTPUT
END_METHOD

METHOD CALL_REQUESTS_EXT
END_METHOD

METHOD CALL_RESETCOMMANDS
END_METHOD

METHOD CALL_RESETOUTPUT
END_METHOD

METHOD CALL_STATEMACHINE
END_METHOD

METHOD CALL_STOP
END_METHOD

METHOD CALL_TMFUNCTIONALITY
END_METHOD

METHOD CALL_ABC
END_METHOD

METHOD CALL_S000_CYCLIC
END_METHOD

METHOD CALL_S001_INIT
END_METHOD

METHOD CALL_S002_READY
END_METHOD

METHOD CALL_S003_HOMING
END_METHOD

METHOD CALL_S010_JOGGING
END_METHOD

METHOD CALL_S011_JOGPOS
END_METHOD

METHOD CALL_S012_JOGNEG
END_METHOD

METHOD CALL_S996_STOP
END_METHOD

METHOD CALL_S998_SERVICE
END_METHOD

METHOD CALL_S999_ERROR
END_METHOD

METHOD CALL_T000_ALLSTATES
END_METHOD

METHOD CALL_T002_READY
END_METHOD

(* ---- _TM_MOTIONCONTROLAXESGROUP.fb ---- *)
FUNCTION_BLOCK _TM_MOTIONCONTROLAXESGROUP EXTENDS _TM_MotionControlBase
VAR_OUTPUT
	XPICKANDPLACEMEMORYLOCK : BOOL;
	EERRORID : L_IE1P_Error;
END_VAR
VAR_IN_OUT
	AXESGROUP : AXES_GROUP_KIN;
	SCCTRLAGBC : scCtrl_AGBC;
	XRESETERROR : BOOL;
	XREGULATORONALL : BOOL;
	XPATHSTOP : BOOL;
	XPATHHALT : BOOL;
	XSTOPALL : BOOL;
	SCPAR : _scPar_TM_MotionControlAGBC;
	SCSTATUSAGBC : scStatus_AGBC;
	XERROR : BOOL;
	XWARNING : BOOL;
	ASCERRORINFO : ARRAY [1..18] OF L_TT1P_scErrorInfo;
	XAXESENABLED : BOOL;
	XAXESGROUPENABLED : BOOL;
	XDONE : BOOL;
	XBUSY : BOOL;
END_VAR
VAR
	XSTOPALL_INT : BOOL;
	IFORCNT : INT;
	DWTEMP : DWORD;
	XABCCTRLREQACTIVE_SAVE : BOOL;
	XRTRIGAGBCJOGGINGINFO : BOOL;
	DWREQUESTSAGBCJOGGINGINFO : DWORD;
	DWREQUESTSAGBCJOGGINGINFO_OLD : DWORD;
	XRTRIGAGBCMOVEINFO : BOOL;
	DWREQUESTSAGBCMOVEINFO : DWORD;
	DWREQUESTSAGBCMOVEINFO_OLD : DWORD;
	XRTRIGAGBCHOMESTOPHALTINFO : BOOL;
	DWREQUESTSAGBCHOMESTOPHALTINFO : DWORD;
	DWREQUESTSAGBCHOMESTOPHALTINFO_OLD : DWORD;
	XRTRIGCTRLABCXSTOP : BOOL;
	DWREQUESTSCTRLABCXSTOP : DWORD;
	DWREQUESTSCTRLABCXSTOP_OLD : DWORD;
	XRTRIGCTRLABCXHALT : BOOL;
	DWREQUESTSCTRLABCXHALT : DWORD;
	DWREQUESTSCTRLABCXHALT_OLD : DWORD;
	XRTRIGCTRLABCXJOGPOS : BOOL;
	DWREQUESTSCTRLABCXJOGPOS : DWORD;
	DWREQUESTSCTRLABCXJOGPOS_OLD : DWORD;
	XRTRIGCTRLABCXJOGNEG : BOOL;
	DWREQUESTSCTRLABCXJOGNEG : DWORD;
	DWREQUESTSCTRLABCXJOGNEG_OLD : DWORD;
	XRTRIGCTRLABCXMOVEVELEXECUTE : BOOL;
	DWREQUESTSCTRLABCXMOVEVELEXECUTE : DWORD;
	DWREQUESTSCTRLABCXMOVEVELEXECUTE_OLD : DWORD;
	XRTRIGCTRLABCXMOVEABSEXECUTE : BOOL;
	DWREQUESTSCTRLABCXMOVEABSEXECUTE : DWORD;
	DWREQUESTSCTRLABCXMOVEABSEXECUTE_OLD : DWORD;
	XRTRIGCTRLABCXMOVERELEXECUTE : BOOL;
	DWREQUESTSCTRLABCXMOVERELEXECUTE : DWORD;
	DWREQUESTSCTRLABCXMOVERELEXECUTE_OLD : DWORD;
	XRTRIGCTRLABCXHOMEEXECUTE : BOOL;
	DWREQUESTSCTRLABCXHOMEEXECUTE : DWORD;
	DWREQUESTSCTRLABCXHOMEEXECUTE_OLD : DWORD;
	XRTRIGCTRLABCXREGULATORON : BOOL;
	DWREQUESTSCTRLABCXREGULATORON : DWORD;
	DWREQUESTSCTRLABCXREGULATORON_OLD : DWORD;
	XERROR_CONCURRENTPICKANDPLACE : BOOL;
	XEXECUTEHALT : BOOL;
	XEXECUTEHALT_OLD : BOOL;
	LRPATHHALTDEC : LREAL;
	LRPATHHALTJERK : LREAL;
	XHALTBUSY : BOOL;
	XHALTDONE : BOOL;
	XHALTCOMANDABROTED : BOOL;
	XEXECUTESTOP : BOOL;
	LRPATHSTOPDEC : LREAL;
	LRPATHSTOPJERK : LREAL;
	XSTOPBUSY : BOOL;
	XSTOPDONE : BOOL;
	XSTOPCOMANDABROTED : BOOL;
	WPATHSTOPSTEPPER : WORD;
	XSTOPALLBUSY : BOOL;
	XSTOPALLDONE : BOOL;
	XSTOPALLCOMANDABROTED : BOOL;
	XTEMPSTOPBUSY : BOOL;
	XTEMPSTOPDONE : BOOL;
	XACCDECSYNC_INT : BOOL;
	XSYNCHRONISED_INT : BOOL;
	XSTOPTRANSITIONLOCK_INT : BOOL;
	XAGBCGROUPSTOPEXECUTE : BOOL;
	XAGBCGROUPSTOPEXECUTEATSYNCOUT : BOOL;
	LRAGBCPATHSTOPDEC : LREAL;
	LRAGBCPATHSTOPJERK : LREAL;
	AGBC : L_MC4P_AxesGroupBasicControl;
	PPARAGBC : POINTER TO _scPar_TM_MotionControlAGBC;
END_VAR
END_FUNCTION_BLOCK

METHOD CALL_ABCCTRLREQACTIVE : BOOL
END_METHOD

METHOD CALL_ABCGENERALSETTINGS
END_METHOD

METHOD CALL_ALLOCPOINTADR
END_METHOD

METHOD CALL_CHECKREQUESTS_ASCCTRLABC
END_METHOD

METHOD CALL_CHECKREQUESTS_SCCTRLAGBC
END_METHOD

METHOD CALL_ERRORHANDLER
END_METHOD

METHOD CALL_ERRORHANDLER_SCERRORINFO
END_METHOD

METHOD CALL_FBMETHODS
END_METHOD

METHOD CALL_FIRSTCYCLE
END_METHOD

METHOD CALL_INITROUTINE
END_METHOD

METHOD CALL_INTERNALCTRL
END_METHOD

METHOD CALL_OUTPUT
END_METHOD

METHOD CALL_REQUESTS_EXT
END_METHOD

METHOD CALL_REQUESTS_ASCCTRLABC
END_METHOD

METHOD CALL_REQUESTS_SCCTRLAGBC
END_METHOD

METHOD CALL_RESETCOMMANDS
END_METHOD

METHOD CALL_RESETOUTPUT
END_METHOD

METHOD CALL_STOP
END_METHOD

METHOD CALL_TMFUNCTIONALITY
END_METHOD

METHOD CALL_AGBC
END_METHOD

METHOD CALL_AGBC_INPUT_ATSERVICE
END_METHOD

METHOD CALL_AGBC_INPUT
END_METHOD

METHOD CALL_PATHSTOPHANDLER
END_METHOD

METHOD CALL_S000_CYCLIC
END_METHOD

METHOD CALL_S001_INIT
END_METHOD

METHOD CALL_S002_READY
END_METHOD

METHOD CALL_S996_STOP
END_METHOD

METHOD CALL_S998_SERVICE
END_METHOD

METHOD CALL_S999_ERROR
END_METHOD

METHOD CALL_T000_ALLSTATES
END_METHOD

(* ---- _TM_MOTIONCONTROLBASE.fb ---- *)
FUNCTION_BLOCK _TM_MOTIONCONTROLBASE EXTENDS _TM_Base
VAR_OUTPUT
	ETMSTATE : L_TT1P_States;
END_VAR
VAR_IN_OUT
	XENABLEINTERNALCONTROL : BOOL;
	XENABLE : BOOL;
	XINTERNALCONTROLACTIVE : BOOL;
END_VAR
VAR
	XSTATEENTRY : BOOL;
	XABCCTRLREQACTIVE : BOOL;
	XTMREQACTIVE : BOOL;
	XTMSTOP : BOOL;
	XINTERNALCONTROL : BOOL;
	XENABLE_INT : BOOL;
	XRESETERROR_INT : BOOL;
	XREGULATORON_INT : BOOL;
	XSTOP_INT : BOOL;
	XHALT_INT : BOOL;
	XHALT_OLD : BOOL;
	SCPARMOTIONCONTROL_INT : _scPar_TM_MotionControl;
	ETMSTATE_OLD : L_TT1P_States;
	REQUESTSINFO : DWORD;
	REQUESTSINFO_OLD : DWORD;
	DWRTRIG : DWORD;
	XNEWREQUEST : BOOL;
	XREQUEST_FTRIG : BOOL;
	DWFTRIG : DWORD;
	BYINBITNO : BYTE;
	XTMWARNING_INT : BOOL;
	XTMERROR_INT : BOOL;
	ETMERRORID_INT : L_IE1P_Error;
	XERROR_FIRST : BOOL;
	EERRORID_FIRST : L_IE1P_Error;
	XRESETERROR_RTRIG : BOOL;
	XRESETOUTPUTDONE : BOOL;
	ETMSTATE_INT : L_TT1P_States;
	XBUSY_INT : BOOL;
	XDONE_INT : BOOL;
	XSWITCHTOSTOP : BOOL;
	XDONENEXTCYCLE_INT : BOOL := TRUE;
	XISHOMED_INT : BOOL;
	LWTCHECKSUM : LWORD;
	XFIRSTCYCLE : BOOL := TRUE;
	ICNTRESETERROR : INT := 10;
	XINITDONE : BOOL;
	IINITSTATE : INT;
	PBOOL : POINTER TO BOOL;
	PBYTE : POINTER TO BYTE;
	PINT : POINTER TO INT;
	PDINT : POINTER TO DINT;
	PUINT : POINTER TO UINT;
	PSINT : POINTER TO SINT;
	PWORD : POINTER TO WORD;
	PDWORD : POINTER TO DWORD;
	PREAL : POINTER TO REAL;
	PLREAL : POINTER TO LREAL;
	PSTRING : POINTER TO STRING;
	DIFRAME : DINT;
	DIFRAMEPAR : DINT;
	C_IJOGGING : INT := 1;
END_VAR
END_FUNCTION_BLOCK

METHOD CALL_ABCCTRLREQACTIVE : BOOL
END_METHOD

METHOD CALL_ABCGENERALSETTINGS
END_METHOD

METHOD CALL_ALLOCPOINTADR
END_METHOD

METHOD CALL_CHECKREQUESTS
END_METHOD

METHOD CALL_CTRLREQACTIVE : BOOL
END_METHOD

METHOD CALL_ERRORHANDLER
END_METHOD

METHOD CALL_FBMETHODS
END_METHOD

METHOD CALL_FIRSTCYCLE
END_METHOD

METHOD CALL_INITDONE
END_METHOD

METHOD CALL_INITROUTINE
END_METHOD

METHOD CALL_INTERNALCTRL
END_METHOD

METHOD CALL_OUTPUT
END_METHOD

METHOD CALL_REQUESTS_EXT
END_METHOD

METHOD CALL_RESETCOMMANDS
END_METHOD

METHOD CALL_RESETOUTPUT
END_METHOD

METHOD CALL_RESETWARNINGS
END_METHOD

METHOD CALL_STATEMACHINE
END_METHOD

METHOD CALL_STOP
END_METHOD

METHOD CALL_TMFUNCTIONALITY
END_METHOD

METHOD CALL_ABC
END_METHOD

METHOD CALL_S000_CYCLIC
END_METHOD

METHOD CALL_S001_INIT
END_METHOD

METHOD CALL_S002_READY
END_METHOD

METHOD CALL_S996_STOP
END_METHOD

METHOD CALL_S998_SERVICE
END_METHOD

METHOD CALL_S999_ERROR
END_METHOD

METHOD CALL_T000_ALLSTATES
END_METHOD

METHOD CALL_T002_READY
END_METHOD

(* ---- _TM_PICKANDPLACEBASE.fb ---- *)
FUNCTION_BLOCK _TM_PICKANDPLACEBASE EXTENDS _TM_MotionControlAxesGroup
VAR_OUTPUT
	PAP : POINTER TO _scAP_TM_PickAndPlaceHigh;
	PSF : POINTER TO _scSF_TM_PickAndPlaceHigh;
END_VAR
VAR_IN_OUT
	FB_EXTERNALMEMORY : L_MC4P_PickAndPlaceMemory;
	SCACCESSPOINTS : _scAP_TM_PickAndPlaceBase;
	XEXECUTEPICKANDPLACE : BOOL;
	XPATHINTERRUPT : BOOL;
	XGROUPHOMEEXECUTE : BOOL;
	AXHOMEABSSWITCH : ARRAY [1..12] OF BOOL;
	XGROUPENABLEHWLIMIT : BOOL;
	AXHWLIMITPOS : ARRAY [1..18] OF BOOL;
	AXHWLIMITNEG : ARRAY [1..18] OF BOOL;
	ESELECTAXIS : IDENT_IN_GROUP_REF;
	XJOGPOS : BOOL;
	XJOGNEG : BOOL;
	XABORT : BOOL;
	LROVERRIDE : LREAL;
	SCSIGNALFLOW : _scSF_TM_PickAndPlaceBase;
	XAXESGROUPHOMED : BOOL;
	XACTIVE : BOOL;
	XHWLIMITSWITCHACTIVE : BOOL;
	XSWLIMITSWITCHACTIVE : BOOL;
	AXHWLIMITSWITCHNEG : ARRAY [1..18] OF BOOL;
	AXHWLIMITSWITCHPOS : ARRAY [1..18] OF BOOL;
	AXSWLIMITSWITCHENABLE : ARRAY [1..18] OF BOOL;
	AXSWLIMITSWITCHACTIVE : ARRAY [1..18] OF BOOL;
	XINPOSITION : BOOL;
	XPATHHOLD : BOOL;
	XGRIPPERCTRLACTIVE : BOOL;
	XPULSEGRIPPER : BOOL;
	LRSETPATHVELOUT : LREAL;
	LRPATHPREPARATIONTIME : LREAL;
	LRPRECALCPROFILETIME : LREAL;
	ALRACTAXISPOS : ARRAY [1..18] OF LREAL;
	ALRACTAXISVEL : ARRAY [1..18] OF LREAL;
	IPROFILEPOINTPASSED : INT;
END_VAR
VAR
	PPARBASE : POINTER TO _scPar_TM_PickAndPlaceBase;
	XEXECUTEPICKANDPLACE_INT : BOOL;
	XPATHINTERRUPT_INT : BOOL;
	XGROUPHOMEEXECUTE_INT : BOOL;
	AXHOMEABSSWITCH_INT : ARRAY [1..12] OF BOOL;
	LRSETPATHVELOUT_INT : LREAL;
	XGROUPENABLEHWLIMIT_INT : BOOL;
	AXHWLIMITPOS_INT : ARRAY [1..18] OF BOOL;
	AXHWLIMITNEG_INT : ARRAY [1..18] OF BOOL;
	XABORT_INT : BOOL;
	LROVERRIDE_INT : LREAL;
	ESELECTAXIS_INT : IDENT_IN_GROUP_REF;
	XJOGPOS_INT : BOOL;
	XJOGNEG_INT : BOOL;
	XENABLEPOSINWINDOW_INT : BOOL;
	XINPOSITION_INT : BOOL;
	LRHOMEPOSITION_INT : LREAL;
	SCHOMEEXTPARAMETER_INT : L_MC1P.L_MC1P_HomeParameter;
	SCHOMEEXTTP_INT : L_MC1P.MC_TRIGGER_REF;
	EHOMINGORDER_INT : L_MC4P.L_MC4P_HomingOrder;
	XABORT_OLD : BOOL;
	XABORT_LOCK : BOOL;
	IDX1 : INT;
	ITMP : INT;
	LRTMP : LREAL;
	LRTMP1 : LREAL;
	LRTMP2 : LREAL;
	LRTMP3 : LREAL;
	TTMP : TIME;
	WID : WORD;
	XPROFILERECEIVEDGAPS : BOOL;
	XPATHINTERRUPTACTIVE : BOOL;
	XPREPARINGPATH_INT : BOOL;
	ECOORDSYSTEMP1 : L_MC4P_CoordSystem := L_MC4P_CoordSystem.MCS;
	XINPOSITIONHOLDSETPOS : BOOL;
	LRTASKCYCLE : LREAL := 0.001;
	LRSTARTXPOS : LREAL;
	LRSTARTYPOS : LREAL;
	LRSTARTZPOS : LREAL;
	LRSTARTAUX1POS : LREAL;
	XOVERRIDEATMOVEPPACTIVE : BOOL;
	XOVERRIDEOUTATMOVEPP : BOOL;
	LROVERRIDEOUTATMOVEPP : LREAL;
	LROVERRIDEFADINGTIMEATMOVEPP : LREAL;
	XWARNINGSELECTEDAXISNOTSUPPORTED : BOOL;
	XWARNINGXSWMAX : BOOL;
	XWARNINGYSWMAX : BOOL;
	XWARNINGZSWMAX : BOOL;
	XWARNINGAUX1SWMAX : BOOL;
	XERRORINVALIDPROFILE : BOOL;
	XERROR_INVALIDCOORDSYSTEM : BOOL;
	XWARNINGAXESGROUPNOTENABLED : BOOL;
	XWARNINGSEMAMOVEFBNOTFREE : BOOL;
	LRGRIPPERCLOSINGTIME_INT : LREAL;
	LRORFADINGTIME_INT : LREAL;
	XLOADORFADINGTIME_INT : BOOL;
	LROVERRIDEFADINGTIME_INT : LREAL;
	LRSETFBOROVERRIDE_INT : LREAL;
	_XLIMITDYNAMICS_ENABLE : BOOL;
	_XPP_ENABLE : BOOL;
	_XPP_ENABLE_OLD : BOOL;
	_XPP_ABORT : BOOL;
	_XPP_EXECUTEPICKANDPLACE : BOOL;
	_LRPP_STARTBLENDINGRADIUS : LREAL;
	_XPP_ERROR : BOOL;
	_EPP_ERRORID : L_IE1P_Error;
	_XPP_BUSY : BOOL;
	_XPP_DONE : BOOL;
	_XPP_COMMANDABORTED : BOOL;
	_XPP_PROFILEINPREPARATION : BOOL;
	_XPP_MOVEPPACTIVE : BOOL;
	_XPP_PATHHOLD : BOOL;
	_IPP_PROFILEPOINTPASSED : INT;
	_IPP_TARGETPROFILEPOINT : INT;
	_ALRPP_TARGETPOSITION : ARRAY [1..12] OF LREAL;
	_EPP_SETSEGMENTTYPEOUT : L_MC4P_SegmentType;
	_BYPP_NUMOFPOINTSINPROFILE : BYTE;
	_BYPP_NUMOFHALTINPROFILE : BYTE;
	_LRPP_PATHPREPARATIONTIME : LREAL;
	_LRPP_PROFILERESTTIME : LREAL;
	_LRPP_PRECALCPROFILETIME : LREAL;
	_XPP_TIMEVALID : BOOL;
	_LRPP_INTERRUPTPATHACC : LREAL;
	_XPP_PATHINTERRUPTOUT : BOOL;
	_XPP_PATHINTERRUPTOUT_OLD : BOOL;
	MP00_LWTCHECKSUM : LWORD;
	MP20_PAMOVELINEARABSOLUTE : POINTER TO ARRAY [1..10] OF L_MC4P_MoveLinearAbsolute_Internal;
	MP21_PAMOVELINEARABSOLUTE : POINTER TO ARRAY [1..10] OF L_MC4P_MoveLinearAbsolute_Internal;
	MP22_PAMOVELINEARABSOLUTE : POINTER TO ARRAY [1..10] OF L_MC4P_MoveLinearAbsolute_Internal;
	MP23_PAMOVELINEARABSOLUTE : POINTER TO ARRAY [1..10] OF L_MC4P_MoveLinearAbsolute_Internal;
	XSEMAMOVEFBS_LOCK : BOOL;
	FB_LIMITDYNAMICSMAINAXES : L_MC4P_LimitDynamicsMainAxes;
	FB_LIMITDYNAMICSAUXAXES : L_MC4P_LimitDynamicsAuxAxes;
	AFB_HWLIMITAXIS : ARRAY [1..13] OF L_MC1P_HWLimitSwitchInterface;
	AFB_INPOSITION : ARRAY [1..6] OF L_TT1P_InPosition;
	FB_SETOVERRIDE : L_MC4P_GroupSetOverride;
	XVISUHOMEABSSWITCH : BOOL;
	STVISUSELECTAXIS : STRING := 'AxisX';
	EVISUSELECTAXIS : IDENT_IN_GROUP_REF := IDENT_IN_GROUP_REF.X;
	EVISUHOMESELECTAXIS : IDENT_IN_GROUP_REF := IDENT_IN_GROUP_REF.A1;
	EVISUHOMESELECTAXIS_OLD : IDENT_IN_GROUP_REF;
	EVISUSELECTAXIS_OLD : L_MC4P.IDENT_IN_GROUP_REF;
	DIFRAME_OLD : DINT;
	LWACTIVELIMITS_MAN : LWORD;
	DWACTIVELIMITS_0_MAN : DWORD;
	DWACTIVELIMITS_1_MAN : DWORD;
	C_BYMAXTARGETPOINTS : BYTE := 10;
END_VAR
END_FUNCTION_BLOCK

METHOD CALL_ALLOCPOINTADR
END_METHOD

METHOD CALL_ERRORHANDLER
END_METHOD

METHOD CALL_FBMETHODS
END_METHOD

METHOD CALL_FB_HWLIMITAXISA
END_METHOD

METHOD CALL_FB_HWLIMITAXISA1
END_METHOD

METHOD CALL_FB_HWLIMITAXISA2
END_METHOD

METHOD CALL_FB_HWLIMITAXISA3
END_METHOD

METHOD CALL_FB_HWLIMITAXISA4
END_METHOD

METHOD CALL_FB_HWLIMITAXISA5
END_METHOD

METHOD CALL_FB_HWLIMITAXISA6
END_METHOD

METHOD CALL_FB_HWLIMITAXISAUX1
END_METHOD

METHOD CALL_FB_HWLIMITAXISB
END_METHOD

METHOD CALL_FB_HWLIMITAXISC
END_METHOD

METHOD CALL_FB_HWLIMITAXISX
END_METHOD

METHOD CALL_FB_HWLIMITAXISY
END_METHOD

METHOD CALL_FB_HWLIMITAXISZ
END_METHOD

METHOD CALL_FB_LIMITDYNAMICSAUXAXES
END_METHOD

METHOD CALL_FB_LIMITDYNAMICSAUXAXES_INPUT
END_METHOD

METHOD CALL_FB_LIMITDYNAMICSMAINAXES
END_METHOD

METHOD CALL_FB_LIMITDYNAMICSMAINAXES_INPUT
END_METHOD

METHOD CALL_FB_OVERRIDE
END_METHOD

METHOD CALL_FB_OVERRIDECONTROL
END_METHOD

METHOD CALL_FB_OVERRIDE_INPUT
END_METHOD

METHOD CALL_FM_MOVEPICKANDPLACE
END_METHOD

METHOD CALL_FM_MOVEPICKANDPLACE_INTPUT
END_METHOD

METHOD CALL_FIRSTCYCLE
END_METHOD

METHOD CALL_INITCHECKINTERMEDIANTEMOVELINABS
END_METHOD

METHOD CALL_INITDONE
END_METHOD

METHOD CALL_INITROUTINE
END_METHOD

METHOD CALL_INTERNALCTRL
END_METHOD

METHOD CALL_MC_GROUPREADACTUALPOSITION
END_METHOD

METHOD CALL_OUTPUT
END_METHOD

METHOD CALL_OUTPUT_SF
END_METHOD

METHOD CALL_PPABORT
END_METHOD

METHOD CALL_REQUESTS_EXT
END_METHOD

METHOD CALL_RESETCOMMANDS
END_METHOD

METHOD CALL_RESETOUTPUT
END_METHOD

METHOD CALL_RESETWARNINGS
END_METHOD

METHOD CALL_SEMAMOVEFB_RELEASE
END_METHOD

METHOD CALL_STATEMACHINE
END_METHOD

METHOD CALL_VISUCTRL
END_METHOD

METHOD CALL_AFB_INPOSITION
END_METHOD

METHOD FUN_GETPATHINTERRUPTORFEEDINGTIME
END_METHOD

METHOD CALL_AGBC_INPUT_ATSERVICE
END_METHOD

METHOD FUN_AXISINPOSITION
VAR_IN_OUT
	PAXIS : POINTER TO AXIS_REF;
	FB_INPOSITION : L_TT1P_InPosition;
	XINPOSITION : BOOL;
END_VAR
END_METHOD

METHOD CALL_S000_CYCLIC
END_METHOD

METHOD CALL_S002_READY
END_METHOD

METHOD CALL_S003_HOMING
END_METHOD

METHOD CALL_S112_PREPARING_PATH
END_METHOD

METHOD CALL_S114_MOVE_PP
END_METHOD

METHOD CALL_S117_PATH_INTERRUPT
END_METHOD

METHOD CALL_S150_JOGGING_X
END_METHOD

METHOD CALL_S151_JOGGING_Y
END_METHOD

METHOD CALL_S152_JOGGING_Z
END_METHOD

METHOD CALL_S153_JOGGING_A
END_METHOD

METHOD CALL_S154_JOGGING_B
END_METHOD

METHOD CALL_S155_JOGGING_C
END_METHOD

METHOD CALL_S156_JOGGING_A1
END_METHOD

METHOD CALL_S157_JOGGING_A2
END_METHOD

METHOD CALL_S158_JOGGING_A3
END_METHOD

METHOD CALL_S159_JOGGING_A4
END_METHOD

METHOD CALL_S160_JOGGING_A5
END_METHOD

METHOD CALL_S161_JOGGING_A6
END_METHOD

METHOD CALL_S162_JOGGING_AUX1
END_METHOD

METHOD CALL_S996_STOP
END_METHOD

METHOD CALL_S999_ERROR
END_METHOD

METHOD CALL_T002_READY
END_METHOD

METHOD CALL_TXX_JOGGINGSELECTAXIS
END_METHOD

(* ---- _TM_PICKANDPLACEBASEEXTENSION.fb ---- *)
FUNCTION_BLOCK _TM_PICKANDPLACEBASEEXTENSION EXTENDS _TM_PickAndPlaceBase
VAR_OUTPUT
	PPAR : POINTER TO _scPar_TM_PickAndPlaceBaseExtension;
END_VAR
VAR
	SCPAR_INT : _scPar_TM_PickAndPlaceBaseExtension;
	FM_MOVEPICKANDPLACE : L_MB1P_MovePickAndPlaceElliptical;
END_VAR
END_FUNCTION_BLOCK

METHOD CALL_ALLOCPOINTADR
END_METHOD

METHOD CALL_FM_MOVEPICKANDPLACE
END_METHOD

METHOD CALL_FM_MOVEPICKANDPLACE_INTPUT
END_METHOD

METHOD CALL_INTERNALCTRL
END_METHOD

METHOD CALL_PPABORT
END_METHOD

METHOD CALL_RESETCOMMANDS
END_METHOD

METHOD CALL_S112_PREPARING_PATH
END_METHOD

(* ---- _TM_PICKANDPLACEHIGH.fb ---- *)
FUNCTION_BLOCK _TM_PICKANDPLACEHIGH EXTENDS _TM_PickAndPlaceState
VAR_IN_OUT
	XADDPROFILE : BOOL;
	ISETPROFILENOOUT : INT;
	XPROFILEINPREPARATION : BOOL;
END_VAR
VAR
	XADDPROFILE_INT : BOOL;
	XENDOFPROFILE : BOOL;
	_XPP_ENDOFPROFILE : BOOL;
	_IPP_SETPROFILENOOUT : INT;
	_XPP_WARNING : BOOL;
	FM_MOVEPICKANDPLACE : L_TF1P_AddProfilePickAndPlace;
END_VAR
END_FUNCTION_BLOCK

METHOD CALL_ERRORHANDLER
END_METHOD

METHOD CALL_FM_MOVEPICKANDPLACE
END_METHOD

METHOD CALL_FM_MOVEPICKANDPLACE_INTPUT
END_METHOD

METHOD CALL_INTERNALCTRL
END_METHOD

METHOD CALL_OUTPUT
END_METHOD

METHOD CALL_OUTPUT_SF
END_METHOD

METHOD CALL_S114_MOVE_PP
END_METHOD

(* ---- _TM_PICKANDPLACESTATE.fb ---- *)
FUNCTION_BLOCK _TM_PICKANDPLACESTATE EXTENDS _TM_PickAndPlaceBase
VAR_OUTPUT
	PPAR : POINTER TO _scPar_TM_PickAndPlaceHigh;
END_VAR
VAR_IN_OUT
	XACKPATHHALT : BOOL;
END_VAR
VAR
	SCPAR_INT : _scPar_TM_PickAndPlaceHigh;
	XACKPATHHALT_INT : BOOL;
	IFORCNT2 : INT;
	ICNTENABLEMOVELINABS : INT;
	BYACKPATHSTOPCNT : BYTE := 0;
	AXHALT_INT : ARRAY [0..10] OF BOOL;
	ARVISPOINTLINES : ARRAY [1..4] OF L_TT1P_scProfilePar;
	IVISUTABLESETPOS : INT := 0;
	IVISUTABLESETPOS_OLD : INT := 0;
	IVISUTABLEMAXPOS : INT := 7;
	XVISPOINTMIN : BOOL;
	XVISPOINTMAX : BOOL;
	XVISUSETPOSUP : BOOL;
	XVISUSETPOSDOWN : BOOL;
	XVISUSETPOSUP_OLD : BOOL;
	XVISUSETPOSDOWN_OLD : BOOL;
	XSCROLBUTTENACTIVE : BOOL;
	TSETTIME : TIME := TIME#400ms;
	TON_SCROLBUTTEN : TON;
END_VAR
END_FUNCTION_BLOCK

METHOD CALL_ALLOCPOINTADR
END_METHOD

METHOD CALL_INITROUTINE
END_METHOD

METHOD CALL_INTERNALCTRL
END_METHOD

METHOD CALL_VIS_TON_SCROLBUTTEN
END_METHOD

METHOD CALL_VISUCTRL
END_METHOD

METHOD CALL_VISUTABCTRL
END_METHOD

METHOD CALL_VISUUPDATETAB
END_METHOD

METHOD CALL_S112_PREPARING_PATH
END_METHOD

(* ---- _TM_PICKANDPLACESTATEEXTENSION.fb ---- *)
FUNCTION_BLOCK _TM_PICKANDPLACESTATEEXTENSION EXTENDS _TM_PickAndPlaceState
VAR
	FM_MOVEPICKANDPLACE : L_MB1P_MovePickAndPlaceState;
END_VAR
END_FUNCTION_BLOCK

METHOD CALL_FM_MOVEPICKANDPLACE
END_METHOD

METHOD CALL_FM_MOVEPICKANDPLACE_INTPUT
END_METHOD

METHOD CALL_OUTPUT_SF
END_METHOD

METHOD CALL_PPABORT
END_METHOD

(* ---- _TM_REGISTERCONTROLBASE.fb ---- *)
FUNCTION_BLOCK _TM_REGISTERCONTROLBASE EXTENDS _TM_ElectricalShaftPosHigh
VAR_OUTPUT
	PPARRC : POINTER TO _scPar_TM_RegisterControlHigh;
	PSFRC : POINTER TO _scSF_TM_RegisterControlHigh;
	PAPRC : POINTER TO _scAP_TM_RegisterControlHigh;
END_VAR
VAR_IN_OUT
	XMARKRECEIVE : BOOL;
	LRACTMARKPOSIN : LREAL;
	LRCYCPOSEXTENCODER : LREAL;
	XLOADREGPOS : BOOL;
	LRLOADREGPOS : LREAL;
	SCSIGNALFLOWRC : _scSF_TM_RegisterControlBase;
	LRSETREGPOSOUT : LREAL;
	LRMARKSENSORPOS : LREAL;
	LRACTMARKERROR : LREAL;
	LRACTMARKDIST : LREAL;
	XMARKRECEIVED : BOOL;
	LRREGMARKPOS : LREAL;
	XCORRACTIVE : BOOL;
	XCORRLIMITED : BOOL;
END_VAR
VAR
	SCPARRC_INT : _scPar_TM_RegisterControlHigh;
	PTPAXISREAL : POINTER TO _AXIS_REF_REAL;
	LRCYCPOSEXTENCODER_INT : LREAL;
	XLOADREGPOS_INT : BOOL;
	LRLOADREGPOS_INT : LREAL;
	LRSENSORTOOLDISTOLD : LREAL;
	LRMARKSENSORPOS_INT : LREAL;
	LRFACTORREGISTERTOMASTER : LREAL;
	LRFACTORMASTERTOREGISTER : LREAL;
	LRFACTORSLAVETOMASTER : LREAL;
	LRFACTORSLAVETOREGISTER : LREAL;
	_LRSYNCDRIVESETGEARBOXPOSOUT : LREAL;
	_LRSYNCDRIVESETTRIMVELOUT : LREAL;
	MP07_LRSETGEARBOXPOSIN : LREAL;
	MP08_LRSETGEARBOXPOSOUT : LREAL;
	MP09_LRSETCLUTCHPOSIN : LREAL;
	_XREGISTERCNTRENABLE : BOOL;
	_XREGISTERCNTRLOADREGPOS : BOOL;
	_LRREGISTERCNTRLOADREGPOS : LREAL;
	_LRREGPOSOUT : LREAL;
	_LRREGMARKPOS : LREAL;
	_XMARKRECEIVED : BOOL;
	_LRACTMARKERROR : LREAL;
	_MARKPOSITIONINREGISTER : LREAL;
	_LRMARKSENSORPOS : LREAL;
	_LRACTMARKDIST : LREAL;
	_XCORRACTIVE : BOOL;
	_XCORRLIMITED : BOOL;
	_LRREGISTERCNTRFACTOR : LREAL;
	_LRREGISTERCNTRDELAYACTSET : LREAL;
	_LRTPAXISDELAYCYCLE : LREAL;
	_LRTPDELAYCYCLESACTPOS : LREAL;
	_DWTPAXISDELAYCYCLE : DWORD;
	_LRRESIDUAL : LREAL;
	MP01_LRSETVELOCITYREGISTER : LREAL;
	MP02_LRINTEGRATORREGPOS : LREAL;
	MP03_LRCORRREGPOS : LREAL;
	MP05_XMARKRECEIVEUNLIMITED : BOOL;
	MP06_LRACTMARKERRORUNLIMITED : LREAL;
	FM_SYNCDRIVEREGCTRL : L_TF1P_SyncDriveRegCtrl;
	FM_REGISTERCONTROL_BASE : L_TF1P_RegisterControlBase;
	FB_GEARBOXREGISTERTOSYNCDRIVE : L_MB1P_GearboxPositionInput;
	FB_DIFFERENTIATEMASTERPOS : L_MC2P_Differentiate;
END_VAR
END_FUNCTION_BLOCK

METHOD CALL_FM_SYNCHRONIZEDDRIVE
END_METHOD

METHOD CALL_FM_SYNCHRONIZEDDRIVE_INPUT
END_METHOD

METHOD CALL_ALLOCPOINTADR
END_METHOD

METHOD CALL_CALCFACTORMASTERTOREGISTER
END_METHOD

METHOD CALL_CALCFACTORREGISTERTOMASTER
END_METHOD

METHOD CALL_CALCFACTORSLAVETOMASTER
END_METHOD

METHOD CALL_CALCFACTORSLAVETOREGISTER
END_METHOD

METHOD CALL_CALCMARKSENSORPOS
END_METHOD

METHOD CALL_CALCMASTEROFFSET
END_METHOD

METHOD CALL_ERRORHANDLER
END_METHOD

METHOD CALL_FBMETHODS
END_METHOD

METHOD CALL_FB_DIFFERENTIATEMASTERPOS
END_METHOD

METHOD CALL_FB_DIFFERENTIATEMASTERPOS_INPUT
END_METHOD

METHOD CALL_FB_GEARBOXREGISTERTOSYNCDRIVE
END_METHOD

METHOD CALL_FB_GEARBOXREGISTERTOSYNCDRIVE_INPUT
END_METHOD

METHOD CALL_FM_REGISTERCONTROL
END_METHOD

METHOD CALL_FM_REGISTERCONTROL_INPUT
END_METHOD

METHOD CALL_INITDONE
END_METHOD

METHOD CALL_INITROUTINE
END_METHOD

METHOD CALL_INIT_FM
END_METHOD

METHOD CALL_INTERNALCTRL
END_METHOD

METHOD CALL_OUTPUT
END_METHOD

METHOD CALL_OUTPUT_SF
END_METHOD

METHOD CALL_RESETOUTPUT
END_METHOD

METHOD CALL_TPCOMPENSATION
END_METHOD

METHOD CALL_S000_CYCLIC
END_METHOD

METHOD CALL_S002_READY
END_METHOD

METHOD CALL_S031_POS_IS_SYNCHRONISED
END_METHOD

METHOD CALL_S036_TRIM_POS_PLUS
END_METHOD

METHOD CALL_S037_TRIM_POS_MINUS
END_METHOD

METHOD CALL_S999_ERROR
END_METHOD

METHOD CALL_T002_READY
END_METHOD

(* ---- _TM_REGISTERCONTROLSTATE.fb ---- *)
FUNCTION_BLOCK _TM_REGISTERCONTROLSTATE EXTENDS _TM_RegisterControlBase
VAR_IN_OUT
	XGEARFACTORCORR : BOOL;
	XGEARFACTORCORRHOLD : BOOL;
	XTEACHMARKWINDOW : BOOL;
	XMARKWINDOWOPEN : BOOL;
	XMARKOUTOFWINDOW : BOOL;
	XMARKNOTDETECTED : BOOL;
	XMARKWINDOWTEACHED : BOOL;
	LRACTGEARFACTORCORR : LREAL;
	XGEARFACTORCORRLIMITED : BOOL;
END_VAR
VAR
	XGEARFACTORCORR_INT : BOOL;
	XGEARFACTORCORRHOLD_INT : BOOL;
	XTEACHMARKWINDOW_INT : BOOL;
	_XMARKWINDOWOPEN : BOOL;
	_XMARKOUTOFWINDOW : BOOL;
	_XMARKNOTDETECTED : BOOL;
	_XMARKWINDOWTEACHED : BOOL;
	_LRACTGEARFACTORCORR : LREAL;
	_XGEARFACTORCORRLIMITED : BOOL;
	MP10_XMARKWINDOWCOMPOUT : BOOL;
	MP11_LRMARKSTACKLENGTH : LREAL;
	MP12_LRMARKSTACKERRORTOTAL : LREAL;
	MP13_XMARKRECEIVEDLIMITED : BOOL;
	MP14_LRACTMARKERRORLIMITED : LREAL;
	FM_REGISTERCONTROL_STATE : L_TF1P_RegisterControlState;
END_VAR
END_FUNCTION_BLOCK

METHOD CALL_ERRORHANDLER
END_METHOD

METHOD CALL_FB_GEARBOXREGISTERTOSYNCDRIVE_INPUT
END_METHOD

METHOD CALL_FM_REGISTERCONTROL
END_METHOD

METHOD CALL_FM_REGISTERCONTROL_INPUT
END_METHOD

METHOD CALL_INTERNALCTRL
END_METHOD

METHOD CALL_OUTPUT
END_METHOD

METHOD CALL_OUTPUT_SF
END_METHOD

METHOD CALL_RESETOUTPUT
END_METHOD

METHOD GET_LRMARKSTACKLENGTH : LREAL
END_METHOD

(* ---- _TM_SMARTTRACKBASE.fb ---- *)
FUNCTION_BLOCK _TM_SMARTTRACKBASE EXTENDS _TM_MotionControl
VAR_OUTPUT
	PPAR : POINTER TO _scPar_TM_SmartTrackHigh;
	PSF : POINTER TO _scSF_TM_SmartTrackHigh;
	PAP : POINTER TO _scAP_TM_SmartTrackHigh;
END_VAR
VAR_IN_OUT
	MASTERAXIS : AXIS_REF;
	SLAVEAXIS : AXIS_REF;
	XSYNCVEL : BOOL;
	XPRODUCTEDGERISE : BOOL;
	LRACTPRODUCTEDGEPOSIN : LREAL;
	XPRODUCTEDGEFALL : BOOL;
	LRACTPOS : LREAL;
	LRACTVEL : LREAL;
	LRACTFOLLOWINGERROR : LREAL;
	XPRODUCTRECEIVED : BOOL;
	LRACTPRODUCTERROR : LREAL;
	LRACTPRODUCTERRORLIMITED : LREAL;
	LRMASTERPOSEDGERISE : LREAL;
	XCORRACTIVE : BOOL;
	XCORRLIMITED : BOOL;
END_VAR
VAR
	XSYNCPOS_INT : BOOL;
	SCPAR_INT : _scPar_TM_SmartTrackHigh;
	XMARKRECEIVE_INT : BOOL;
	XMARKRECEIVEOLD : BOOL;
	XMAXCORRECTIONNEG : BOOL;
	XMAXCORRECTIONPOS : BOOL;
	LRACTMARKERRORLIMITED : LREAL;
	XPRODUCTDETECTED_INT : BOOL;
	BYSTEPPER : BYTE;
	BYERRORSTEPPER : BYTE;
	LRDISTANCETOSTOPPOSITION : LREAL;
	FOLLOWSETVALUES1 : L_MC1P_FollowSetValues;
	CONVAXISVELOCITY1 : L_MC2P_ConvAxisV;
	CLUTCHVELOCITY1 : L_TT1P_ClutchVelocity;
	PHASECORRECTIONVEL : L_T01S_PhaseCorrectionVel;
	TOF_CORSENSOR : TOF;
	TRACKCORRECTIONCORSENSOR : L_T01S_PhaseCorrectionVel;
	FILTERPRODUCTDETECTION1 : L_TT1P_FilterProductDetection;
	CALCPRODUCTERROR1 : L_TT1P_CalcProductError_Advanced;
	L_MC1P_TPLIMITDIFF_0 : L_MC1P_TpLimitDiff;
	CONVERTTPPOSITION : L_TT1P_CalculateTPOnMaterialPos_intern;
	TPCOMPFACTOR : L_MB1P_CalculateTpCompensationFactor;
	RTERROR : R_TRIG;
	LRACTMARKPOSIN_INT : LREAL := 0;
	LRACTMARKPOSINRECALC_INT : LREAL := 0;
	LRSETVELOUT_INT : LREAL;
	LRCORRECTIONVALUE : LREAL;
	LRCORRECTIONUNLIMITED : LREAL;
	XCORRECTIONLIMITED_INT : BOOL;
	LRACTMARKERRORLIMITED_INT : LREAL;
	LRLASTSCANOUT : LREAL := 0;
	LRVELOCITYFACTOR_INT : LREAL;
	LRACTMARKERRORLIM_OUT : LREAL;
	LRACTMARKERROR_OUT : LREAL;
	XMARKRECEIVEFALL_INT : BOOL;
END_VAR
END_FUNCTION_BLOCK

METHOD CALL_ALLOCPOINTADR
END_METHOD

METHOD CALL_CLUTCHVELOCITY
END_METHOD

METHOD CALL_CONVAXISVELOCITY
END_METHOD

METHOD CALL_ERRORCALCULATION
END_METHOD

METHOD CALL_ERRORHANDLER
END_METHOD

METHOD CALL_FBMETHODS
END_METHOD

METHOD CALL_FBS
END_METHOD

METHOD CALL_FIRSTCYCLE
END_METHOD

METHOD CALL_FOLLOWSETVALUES
END_METHOD

METHOD CALL_INITDONE
END_METHOD

METHOD CALL_INITROUTINE
END_METHOD

METHOD CALL_INTERNALCTRL
END_METHOD

METHOD CALL_LIMITCORRECTION
END_METHOD

METHOD CALL_OUTPUT
END_METHOD

METHOD CALL_PARAMETER
END_METHOD

METHOD CALL_REQUESTS_EXT
END_METHOD

METHOD CALL_RESETCOMMANDS
END_METHOD

METHOD CALL_RESETOUTPUTS
END_METHOD

METHOD CALL_STATEMACHINE
END_METHOD

METHOD CALL_TOUCHPROBESOURCE
END_METHOD

METHOD CALL_TRACKCORRECTION
END_METHOD

METHOD CALL_ABC
END_METHOD

METHOD CALL_S000_CYCLIC
END_METHOD

METHOD CALL_S041_VEL_IS_SYNCHRONISED
END_METHOD

METHOD CALL_S052_ACC_DEC
END_METHOD

METHOD CALL_S996_STOP
END_METHOD

METHOD CALL_S999_ERROR
END_METHOD

METHOD CALL_T002_READY
END_METHOD

METHOD CALL_T041_VEL_IS_SYNCHRONISED
END_METHOD

METHOD CALL_T052_ACC_DEC
END_METHOD

(* ---- _TM_SMARTTRACKSTATE.fb ---- *)
FUNCTION_BLOCK _TM_SMARTTRACKSTATE EXTENDS _TM_SmartTrackBase
VAR_IN_OUT
	DATABUSIN : ITF_DataBus;
	DATABUSOUT : ITF_DataBus;
	XCOMMUNICATIONVALID : BOOL;
	XMASTER : BOOL;
	XSLAVE : BOOL;
	BYSMARTTRACKNO : BYTE;
	LRDISTTOOUTFEED : LREAL;
END_VAR
VAR
	IOWNTRACKNUMBERINV : INT;
	FIRSTINITIALISATIONCYCLE : BOOL := TRUE;
	ICOUNT : INT;
	LRDISTANCETOMASTER : LREAL;
	IMAXNUMBEROFTRACKS : INT;
	LRSMARTTRACKLENGTHOLD_INT : LREAL;
	LRSENSORPOSITIONOLD_INT : LREAL;
	XINITDONEOLD : BOOL;
	XPARAMETERCHANGE : BOOL;
	XPARAMETERSLAVES : BOOL;
	IOWNTRACKNUMBER : INT;
	XMODULEINITDONE : BOOL;
	BYINITIALISATIONCOUNTER : BYTE := 0;
	XINITMODULECOMMDONE : BOOL;
	XTESTREF : BOOL := FALSE;
	XMODULEREGISTRATIONCOMPLETE : BOOL;
	XINITIALIZED : BOOL;
	PELEMENT : POINTER TO L_MB1P_ChannelElement;
	PRIGHT : POINTER TO L_MB1P_ChannelElement;
	PLEFT : POINTER TO L_MB1P_ChannelElement;
	PDATA : POINTER TO L_MB1P_ChannelData;
	PDATACONTROL : POINTER TO L_MB1P_ChannelData;
	PDATALEFTMODULE : POINTER TO L_MB1P_ChannelData;
	PLIST : POINTER TO L_MB1P_ListControl;
	XLOCKCOMCHANNEL_INT : BOOL;
	IDX : INT;
	XCOMCTRLENABLE : BOOL;
	_XCOMERROR : BOOL;
	_ECOMERRORID : WORD;
	_XCOMERRORINVALIDMASTERCONTROLMODUL : BOOL;
	XWARNINGCOMMUNICATION : BOOL;
	XERRORCOMMUNICATION : BOOL;
	CAMCORRECTION : ARRAY [0..4] OF L_MC2P_CamDataXYVA;
	CAMGETSLAVEPOSITION : L_MC2P_CamGetSlavePosition;
	CAMREF : L_MC2P_CamRefFromStruct;
	LRCORRECTIONPOS : ARRAY [1..10] OF LREAL;
	CLUTCHVELOCITYOFFSET : L_TT1P_ClutchVelocity;
	R_TRIG : R_TRIG;
	F_TRIG : F_TRIG;
	CORRECTTARGETPOSITION : L_TT1P_CorrectTargetPosition;
	R_TRIG_CALCOFFSETACC : R_TRIG;
	FB_COMCHANNEL : L_MB1P_ComChannelState;
	XRESETERROR_COMIN : BOOL;
	AXCURVEACTIVE : ARRAY [1..10] OF BOOL;
	AXSEGMENTACTIVE : ARRAY [1..10] OF BOOL;
	AXSEGMENTACTIVEOLD : ARRAY [1..10] OF BOOL;
	AXCURVEDONE : ARRAY [1..10] OF BOOL;
	ALREXACTDISTANCESTOCONVEYOR : ARRAY [1..10] OF LREAL;
	ALRACTXPOSITION : ARRAY [1..10] OF LREAL;
	ALRACTYPOSITION : ARRAY [1..10] OF LREAL;
	ALRACTPRODUCTPOS : ARRAY [1..10] OF LREAL;
	ALRACTPRODUCTPOSOUT : ARRAY [1..10] OF LREAL;
	ALRACTYVELOCITY : ARRAY [1..10] OF LREAL;
	ALROLDYPOSITION : ARRAY [1..10] OF LREAL;
	ALRTPERROR : ARRAY [1..10] OF LREAL;
	ALRSWITCHVELDIST : ARRAY [1..10] OF LREAL;
	ALRSWITCHVELOCITYPOSITION : ARRAY [1..10] OF LREAL;
	ALRSETVELOCITYOFFSET : ARRAY [1..10] OF LREAL;
	ALRREMAINMULTIPLEBELTCORR : ARRAY [1..10] OF LREAL;
	ALRV : ARRAY [1..10] OF LREAL;
	ALRV0 : ARRAY [1..10] OF LREAL;
	ALRSETVELOCITYOFFSET1 : ARRAY [1..10] OF LREAL;
	ALRSETVELOCITYOFFSET2 : ARRAY [1..10] OF LREAL;
	AICAMSINSEGMENT : ARRAY [1..10] OF INT;
	AICAMSINSEGMENTOLD : ARRAY [1..10] OF INT;
	ALRALLTRACKJERK : ARRAY [1..10] OF LREAL;
	ALRALLTRACKACC : ARRAY [1..10] OF LREAL;
	ICOUNTER : INT := 1;
	LRCOMBINEDSMARTTRACKLENGTH : LREAL := 0;
	LRNORMEDXPOSITION : LREAL;
	LRNORMEDYPOSITION : LREAL;
	LRACCCLUTCH : LREAL := 1000;
	LRJERKCLUTCH : LREAL := 1000000;
	ICOUNTER2 : INT;
	LRCOMBINEDBELTLENGTH : LREAL;
	ITRACK : INT;
	ICAMDATA : INT;
	XVELOCITYOFFSETFLAG : BOOL := FALSE;
	LRSETVELOCITY : LREAL;
	DWBITMASK : DWORD := 4294967295;
	DWSETBIT : DWORD;
	DWTEST : DWORD;
	LRCAMCORRECTIONVELOCITY_INT : LREAL;
	LRCAMCORRECTIONACC_INT : LREAL;
	LRCAMCORRECTIONJERK_INT : LREAL;
	DWVELOCITYCHANGEBITS : DWORD;
	LRREMAINMULTIPLEBELTCORR_INT : LREAL;
	LRTOTALCORRECTIONVALUE : LREAL;
	LRPRODUCTLENGTH_INT : LREAL;
	LRMULTIPLEBELTCLUTCHTIME : LREAL;
	XMULTIPLEBELTCORRECTIONACTIVE_INT : BOOL;
	LRVELOCITYFACTORMASTER_INT : LREAL;
	LRDISTANCETOCONVEYOR : LREAL;
	I : INT;
	IARRAYOFFSET : INT := 0;
	LRMULTIPLEBELTJERK_INT : LREAL;
	LRPRODUCTTARGET_INT : LREAL;
	LRPRODUCTTARGETCORRECTED : LREAL;
	LROFFSETVELOCITYOLD : LREAL;
	XCAMCORRECTIONINVALID : BOOL;
	LRALLTRACKSYNCDIST_INT : LREAL := 1;
	XJERKACTIVE : BOOL;
	ALRALLTRACKACCTIME : ARRAY [1..10] OF LREAL;
END_VAR
END_FUNCTION_BLOCK

METHOD CALL_CALCOFFSETCLUTCHPARAMETER
END_METHOD

METHOD CALL_CALCULATEACTIVECAMS
END_METHOD

METHOD CALL_CAMDATA
END_METHOD

METHOD CALL_CAMGETSLAVEPOSITION
END_METHOD

METHOD CALL_CLUTCHVELOCITYOFFSET
END_METHOD

METHOD CALL_COMIN_POSBASED
END_METHOD

METHOD CALL_COMOUT_POSBASED
END_METHOD

METHOD CALL_ERRORCALCULATION
END_METHOD

METHOD CALL_ERRORHANDLER
END_METHOD

METHOD CALL_FB_COMCHANNEL
END_METHOD

METHOD CALL_FBS
END_METHOD

METHOD CALL_FOLLOWSETVALUES
END_METHOD

METHOD CALL_INITCAMREFS
END_METHOD

METHOD CALL_INITDONE
END_METHOD

METHOD CALL_INTERNALCTRL
END_METHOD

METHOD CALL_OUTPUT
END_METHOD

METHOD CALL_PARAMETER
END_METHOD

METHOD CALL_PRODUCTPOSITION
END_METHOD

METHOD CALL_SHIFTARRAYS
END_METHOD

METHOD CALL_SHIFTPRODUCTPOSITION
END_METHOD

METHOD CALL_SLAVECORRECTIONVEL_POSBASED
END_METHOD

METHOD CALL_TRACKCORRECTION
END_METHOD

METHOD CALL_S000_CYCLIC
END_METHOD

METHOD CALL_S002_READY
END_METHOD
